(* IEC 61131-3 sources: daoli-st-library/DL_Algo (part 12) *)

(* ---- FB_DL_EtchEndpointTrend.st ---- *)
(*==============================================================================
 * 组件名称 (Component)  : FB_DL_EtchEndpointTrend
 * 所属子库 (Sublibrary) : DL_Algo
 * 前缀     (Prefix)     : FB_DL_
 * 当前版本 (Version)    : 1.0.1
 * 兼容性   (Platform)   : CODESYS 3.5 / TwinCAT 3 / 汇川 InoProShop / Schneider
 *                         Machine Expert；纯 IEC 61131-3（第 3 版），
 *                         仅依赖标准库 TON / ABS / MAX / MIN 与库内
 *                         FB_DL_Differentiator（IN-OUT 注入消费），
 *                         零厂商方言
 * 作者     (Author)     : 道莅代码库 · PLC编程专家（R31）
 * 开源溯源 (Origin)     : 刻蚀终点趋势检测公开工艺语义（行业池主源；
 *                         Measurement 行统计族语义邻接不重复记账），道莅
 *                         clean-room 防御性实现，未复制任何外部源码行
 * 功能描述 (Function)   : 刻蚀终点趋势双判据检测件。学习相采基线（均值与
 *                         噪声窗）；监视相用库内 FB_DL_Differentiator 求变化
 *                         率（IN-OUT 注入，不内联），斜率换算为 单位每分钟；
 *                         双判据：斜率绝对值超阈 且 信号突破噪声窗，持续
 *                         tConf 触发终点并锁存，保持至 bRun 下降显式复位。
 *                         斜率量纲占位说明：fSignal 的工程单位由调用方定义，
 *                         fSlope 与 fSlopeTh 同量纲，单位为 调用方单位每分钟。
 * 依赖表   (Depends)    : FB_DL_Differentiator（微分器，IN-OUT 注入消费，
 *                         本件不内联差分）。
 * 状态机   (States)     : eLearning/eMonitor/eTriggered，CASE 带 ELSE 复位
 *                         回学习相（信息级提示）。
 * 码位     (Codes)      : 16#0002_3033 信息级：信号非有限冻结评估、学习相
 *                                      非有限重启学习、样本不足不出判定
 *                                      （不置 bError）
 *                         16#0002_3034 故障级：确认窗中断判据矛盾（锁存）
 *                         16#0002_3035~0037 保留未启用（码表与实现对齐）
 * 边界防错 (Boundary)   : 1 信号非有限（x<>x 自反判加幅值界）监视相冻结评估、
 *                           学习相清积累重启学习；
 *                         2 学习相样本不足不出判定；
 *                         3 斜率时间差防除零由库内微分器公共钳位承担
 *                           （其 fDt 下限 10 毫秒），本件不做二次除法；
 *                         4 TON 实例每拍无条件刷新；
 *                         5 触发锁存可达解除路径：bRun 下降沿显式复位；
 *                         6 确认窗中途判据消失按判据矛盾锁故障。
 * 修订历史 (Revision)   : 2026-11-18 v1.0.0 首版入库（R31 · 阶段三 · 序 20）
 *                         2026-11-18 v1.0.1 R31 终审修复：先验基线模式补
 *                         uCnt 计数，消除方差分母 1E-30 退化致判据二永假
 *==============================================================================*)

(*------------------------------------------------------------------------------
 * 枚举: E_DL_EndpointState（归属本功能块，同文件发布，全库唯一属主）
 *----------------------------------------------------------------------------*)
TYPE E_DL_EndpointState :
(
    eLearning  := 0,   // 学习相：采基线均值与噪声窗 / Learning, baseline mean and noise window
    eMonitor   := 10,  // 监视相：双判据评估 / Monitor, dual-criteria evaluation
    eTriggered := 20   // 触发相：终点锁存至显式复位 / Triggered, endpoint latched until explicit reset
);
END_TYPE

(*==============================================================================
 * 功能块: FB_DL_EtchEndpointTrend
 * 调用约定: 每个扫描周期无条件调用一次；ioDiff 为调用方持有的库内微分器
 *           实例（IN-OUT 注入），本件驱动其引脚并读取其输出。
 *==============================================================================*)
FUNCTION_BLOCK FB_DL_EtchEndpointTrend
VAR_INPUT
    fSignal   : LREAL := 0.0;         // 工艺信号 [调用方单位] / Process signal [caller unit]
    bRun      : BOOL := FALSE;        // 工步运行（下降沿显式复位）/ Process running, falling edge resets
    fSlopeTh  : REAL := 5.0;          // 斜率判据阈 [调用方单位每分钟] / Slope threshold [caller unit per min]
    fNoiseWin : REAL := 2.0;          // 噪声窗 [调用方单位] / Noise window [caller unit]
    tConf     : TIME := T#3S;         // 触发确认窗时长 [毫秒] / Trigger confirm window [ms]
    fBaseline : LREAL := 0.0;         // 外部先验基线（0 = 无先验走自采）/ External prior baseline, 0 = none
    tLearn    : TIME := T#30S;        // 学习相时长 [毫秒]（可增引脚）/ Learning duration [ms], added pin
    tSample   : TIME := T#500MS;      // 微分器采样周期 [毫秒]（可增引脚）/ Differentiator sample period [ms], added pin
END_VAR
VAR_IN_OUT
    ioDiff    : FB_DL_Differentiator; // 库内微分器实例注入（斜率不内联）/ Library differentiator instance injected
END_VAR
VAR_OUTPUT
    bEndpoint : BOOL;                 // 终点触发锁存输出 / Endpoint trigger latched output
    fSlope    : REAL;                 // 斜率输出 [调用方单位每分钟] / Slope output [caller unit per min]
    eState    : E_DL_EndpointState;   // 判定状态 / Detection state
    bError    : BOOL;                 // 故障标志，与故障级码配对（R45）/ Fault flag paired with fault codes
    uErrorId  : UDINT;                // 错误码，0 = 无错 / Error code, 0 = none
END_VAR
VAR
    tonLearn  : TON;                  // 学习相计时，每拍无条件刷新 / Learning timer, refreshed every scan
    tonConf   : TON;                  // 触发确认窗计时，每拍无条件刷新 / Confirm window timer, refreshed every scan
    fSigR     : REAL;                 // 信号 REAL 域副本 [调用方单位] / Signal REAL copy [caller unit]
    bSigOk    : BOOL;                 // 信号有限有效 / Signal finiteness validity
    fSum      : REAL;                 // 学习相样本和 [调用方单位] / Learning sample sum [caller unit]
    fSumSq    : REAL;                 // 学习相平方和 [平方调用方单位] / Learning sum of squares
    uCnt      : UDINT;                // 学习相样本数 [个] / Learning sample count
    fMean     : REAL;                 // 基线均值 [调用方单位] / Baseline mean [caller unit]
    fNoise    : REAL;                 // 噪声窗实测 [调用方单位] / Measured noise window [caller unit]
    bLearnDone: BOOL;                 // 学习完成标志 / Learning done flag
    bCritSlope: BOOL;                 // 判据一：斜率超阈 / Criterion one, slope over threshold
    bCritNoise: BOOL;                 // 判据二：突破噪声窗 / Criterion two, beyond noise window
    bCritNow  : BOOL;                 // 双判据本拍合取 / Both criteria this scan
    bInWin    : BOOL;                 // 确认窗进行中 / Confirm window in progress
    bPriorUse : BOOL;                 // 先验基线使用标志 / Prior baseline usage flag
    uCodeLatch: UDINT;                // 故障级锁存码 / Latched fault code
END_VAR
VAR CONSTANT
    DL_EET_FIN   : LREAL := 1.0E30;   // LREAL 有限幅值判界 / LREAL finiteness magnitude bound
    DL_EET_FINR  : REAL  := 1.0E30;   // REAL 有限幅值判界 / REAL finiteness magnitude bound
    DL_EET_MIN   : UDINT := 20;       // 学习相最少样本数 [个] / Learning minimum samples
    DL_EET_MIN60 : REAL  := 60.0;     // 每秒到每分钟换算系数 / Per-second to per-minute factor
    DL_EET_EPS   : REAL  := 1.0E-30;  // 样本数防除零容差 / Sample count divide guard
END_VAR

// ---- 段 1｜定时器实例无条件周期刷新（红线：禁入条件分支）----------------------
tonLearn(IN := (eState = eLearning) AND bRun, PT := tLearn);   // 学习计时 / Learning timing
tonConf(IN := bCritNow, PT := tConf);                          // 确认窗计时无条件 / Confirm timing unconditionally

// ---- 段 2｜信号有效性（自反判加幅值界）----------------------------------------
bSigOk := (fSignal = fSignal) AND (ABS(fSignal) < DL_EET_FIN); // 信号有限 / Signal finite
fSigR := LREAL_TO_REAL(fSignal);                               // 信号落 REAL 域 / Signal to REAL domain

// ---- 段 3｜显式复位：bRun 下降沿清全部锁存 ------------------------------------
IF NOT bRun THEN
    bEndpoint := FALSE;                            // 复位清终点锁存 / Reset clears endpoint latch
    IF eState = eTriggered THEN
        eState := eLearning;                       // 触发相复位回学习 / Triggered resets to learning
    END_IF
END_IF

// ---- 段 4｜驱动库内微分器（IN-OUT 注入，输出即变化率 单位每秒）----------------
ioDiff(bEnable := bRun AND bSigOk,                    // 信号无效停微分防伪速率 / Invalid signal stops differentiator
       fIn := fSigR,                                  // 被微分量注入 / Differentiated input injected
       tFiltTime := T#1S,                             // 低通时间常数固定档 / Fixed low-pass constant
       tSampleTime := tSample);                       // 采样周期透传 / Sample period passed
fSlope := ioDiff.fRateOut * DL_EET_MIN60;             // 斜率换算每分钟（量纲占位见头注释）/ Slope per minute

// ---- 段 5｜学习相：采基线均值与噪声窗 ------------------------------------------
IF (eState = eLearning) AND bRun THEN
    IF NOT bSigOk THEN
        fSum := 0.0;                                  // 非有限清积累重启学习（信息级）/ Non-finite restarts learning
        fSumSq := 0.0;                                // 清平方和积累 / Clear sum-of-squares
        uCnt := 0;                                    // 清样本计数 / Clear sample count
        bLearnDone := FALSE;                          // 撤完成标志 / Withdraw done flag
        uErrorId := 16#0002_3033;                     // 信息级：学习重启 / Info: learning restarted
    ELSE
        bPriorUse := (fBaseline <> 0.0) AND (fBaseline = fBaseline)
                 AND (ABS(fBaseline) < DL_EET_FIN);   // 先验基线可用性 / Prior baseline availability
        IF bPriorUse THEN
            fMean := LREAL_TO_REAL(fBaseline);        // 先验均值直接生效 / Prior mean applied directly
            uCnt := uCnt + 1;                         // 先验模式同样计数（方差分母防爆，R28 终审）/ Prior mode counts samples too
        ELSE
            fSum := fSum + fSigR;                     // 自采样本累加 / Self-sample accumulation
            uCnt := uCnt + 1;                         // 样本计数 / Sample count
        END_IF
        fSumSq := fSumSq + fSigR * fSigR;             // 平方和积累（样本方差用）/ Sum of squares accumulation
        IF tonLearn.Q AND (bPriorUse OR (uCnt >= DL_EET_MIN)) THEN
            IF NOT bPriorUse THEN
                fMean := fSum / UDINT_TO_REAL(uCnt);  // 均值收口，分母已验下限 / Mean closed, denominator verified
            END_IF
            fNoise := SQRT(MAX(fSumSq / MAX(UDINT_TO_REAL(uCnt), DL_EET_EPS) - fMean * fMean, 0.0)); // 样本标准差收口（平方和法）/ Sample stddev via sum-of-squares
            bLearnDone := TRUE;                       // 学习完成 / Learning done
            eState := eMonitor;                       // 转监视相 / To monitor
        END_IF
    END_IF
END_IF

// ---- 段 6｜监视相：双判据评估与确认窗 ------------------------------------------
IF (eState = eMonitor) AND bRun THEN
    IF NOT bSigOk OR (NOT ioDiff.bValid) THEN
        bCritSlope := FALSE;                          // 数据无效撤判据一 / Invalid data withdraws criterion one
        bCritNoise := FALSE;                          // 数据无效撤判据二 / Invalid data withdraws criterion two
        uErrorId := 16#0002_3033;                     // 信息级：冻结评估 / Info: evaluation frozen
    ELSIF (uCnt < DL_EET_MIN) AND (NOT bPriorUse) THEN
        bCritSlope := FALSE;                          // 样本不足不出判定 / Insufficient samples, no verdict
        bCritNoise := FALSE;                          // 样本不足不出判定 / Insufficient samples, no verdict
        uErrorId := 16#0002_3033;                     // 信息级：样本不足 / Info: insufficient samples
    ELSE
        bCritSlope := ABS(fSlope) > ABS(fSlopeTh);    // 判据一：斜率超阈 / Slope over threshold
        bCritNoise := ABS(fSigR - fMean) > fNoise;    // 判据二：突破噪声窗 / Beyond noise window
    END_IF
    bCritNow := bCritSlope AND bCritNoise;            // 双判据合取 / Both criteria AND
    bInWin := (tonConf.ET > T#0MS);                   // 确认窗进行中判定 / Confirm window in progress
    IF bInWin AND (NOT bCritNow) THEN
        eState := eLearning;                          // 按判据矛盾复位回学习重采基线 / Contradiction resets to learning
        uCodeLatch := 16#0002_3034;                   // 码位：确认窗中断判据矛盾 / Code: confirm window contradiction
        bError := TRUE;                               // 故障级配对置位（R45）/ Fault flag paired
    ELSIF tonConf.Q THEN
        bEndpoint := TRUE;                            // 确认满终点触发锁存 / Confirmed, endpoint latched
        eState := eTriggered;                         // 转触发相 / To triggered
        bError := FALSE;                              // 清故障标志 / Clear fault flag
        uCodeLatch := 16#0000_0000;                   // 清锁存码 / Clear latched code
    END_IF
END_IF

// ---- 段 7｜错误码装配：故障锁存回放优先，信息级居次 -----------------------------
IF (eState = eLearning) AND bRun AND (uCodeLatch <> 16#0000_0000) THEN
    bError := TRUE;                                   // 故障锁存回放（学习相等待重试）/ Fault latched replay
    uErrorId := uCodeLatch;                           // 锁存码回放 / Latched code replayed
ELSIF NOT bRun THEN
    bError := FALSE;                                  // 撤运行清故障（可达解除）/ Run drop clears fault
    uErrorId := 16#0000_0000;                         // 清码 / Clear code
    uCodeLatch := 16#0000_0000;                       // 清锁存码 / Clear latched code
END_IF
END_FUNCTION_BLOCK

(* ---- FB_DL_EwmaFilter.st ---- *)
(*
  ==================================================================
  组件名 Component  : FB_DL_EwmaFilter
  分类   Category   : DL_Algo
  前缀   Naming     : FB_DL_ ｜ b/n/u/f/t/e/st 类型前缀制（R265）
  码位   Code ID    : 16#0002_373B / 373C（故障级）
  版本   Version    : 1.0.0
  复杂度 Complexity  : 低
  功能   Purpose    : EWMA 指数加权滑动平均 fOut := fOut + α×(fIn − fOut)，α 直接
                      入参（离散统计 / SPC 平滑口径），供调用方直接整定平滑系数。
  开源溯源 Origin    : 公开公式 clean-room，参考公开统计过程控制（SPC）教材的
                      EWMA 定义（分类与公式借鉴，零代码复制），本件实现、闸门与
                      码位 100% 自有。
  许可证 License    : MIT
  参考   Reference  : IEC 61131-3:2013 §6.6 算术运算符；EWMA 递推式 y[k] =
                      y[k−1] + α·(x[k] − y[k−1]) 为公开统计公式
  平台   Platform   : 纯 IEC 61131-3（四则 / 比较），三平台通用
  依赖   Depends    : 仅 Standard.library（无库调用、无定时器）
  分工声明 Split     : FB_DL_LowPassFilter 为连续时间常数口径（α 由 tTf / tDt 派生，
                      一阶 RC 语义）；FB_DL_MovingAverage 为等权滑窗；本件为调用方
                      直接给 α 的统计平滑口径（EWMA / SPC 语义）；三者选型对照进
                      MANUAL_DL_Algo（R216 双向互引）。
  归属 Ownership     : 本件无 TYPE 声明；全部引脚为 IEC 标准原生类型。
  ------------------------------------------------------------------
  边界 Boundary     :
                      一 α 域闸 (0, 1]：fAlpha <= 0 或 > 1 或非有限 → 组态码 373B +
                         出口三件套 + RETURN 结构早退（开区间下界防输出冻结，
                         α = 0 是「禁冻结伪装正常」的组态错误而非合法参数）；
                      二 fIn 非有限（NaN / ±Inf）→ 本拍拒绝更新、保持上拍有效值 +
                         故障码 373C + 三件套（禁污染物进入递推状态）；
                      三 首拍 _bInit → fOut := fIn 首样本直通（禁输出 0 假跳变）；
                      四 bEnable = FALSE 的语义写死（FB33-4 声明行）：本件取「冻结
                         最后有效值」，理由：纯监视滤波不驱动功率级，冻结均值供
                         HMI 连续读数（与 BiquadFilter 的「控制量归零」口径不同，
                         选型时注意）；
                      五 故障码策略（本件无 bReset 引脚，R152 解除路径自证）：组态类
                         与测量类故障码逐拍重算不锁存，解除路径 = 修正组态 / 恢复
                         测点（恒可达）；首因保序由判据顺序保证；
                      六 非有限闸逐个点名（R272）：fAlpha 与 fIn 双双入闸；
                      七 首拍 _bInit 全量初始化（FB50-2）；无定时器 / 无边沿实例，
                         段 0 无刷新对象（R6 标注 N/A）；无全局、无外部变量、无
                         物理地址、无指针。
  错误码 Codes      :
    16#0002_373B【故障级】组态非法（fAlpha ≤ 0 / > 1 / 非有限）
    16#0002_373C【故障级】输入非有限（fIn 为 NaN / ±Inf）或递推结果非有限（后者
                         理论上不可达的兜底分支，与输入坏同码，出口组合不可区分，
                         R90 反证：fOut 保持上拍有效值 + bValid = FALSE 两场景同形）
  码位反证 Note     :
    373B 与 373C 不可合并：两者的处置人不同（组态工程师调 α / 仪表工查测点），
    而两者出口组合不同（组态坏无论 fIn 有限与否恒发 373B），可由场景唯一还原，
    故分立两码（R90）。
  验收 Acceptance   :
    算法已证（脚本）：未跑 ｜ 编译器已证（三平台）：未跑
    V1 α = 1 → 直通 fOut = fIn（逐拍断言）
    V2 α = 0 → 码 373B + 三件套 + 早退（禁冻结伪装正常）
    V3 α = 0.5 阶跃 0 → 100 → 逐拍 50 / 75 / 87.5 收敛，无超调
    V4 fIn = NaN → 保持上拍 fOut + 码 373C + bValid = FALSE
    V5 首拍 → fOut = fIn 首样本直通（禁 0 假跳变）
    V6 bEnable = FALSE → fOut 冻结最后有效值（边界四声明行回归向量）
  修订记录 Revision  :
    2026-11-21  v1.0.0  R63 首版（批 1 · 序号 3）
  ==================================================================
*)
FUNCTION_BLOCK FB_DL_EwmaFilter
VAR_INPUT
    bEnable  : BOOL := TRUE;  // 使能，FALSE 时输出冻结最后有效值（边界四）/ the enable, false freezes the last valid output
    fIn      : LREAL := 0.0;  // 输入量 [工程单位]，必须有限 / the input value, must be finite
    fAlpha   : LREAL := 0.2;  // 平滑系数 [−]，合法域 (0, 1] 开区间下界 / the smoothing factor inside the half open domain from zero exclusive to one
END_VAR
VAR_OUTPUT
    fOut     : LREAL := 0.0;           // 滤波输出 [工程单位] / the filtered output
    bValid   : BOOL := FALSE;          // 输出可用（使能 + 无故障 + 首样本已收）[-] / the output is usable
    eErr     : UDINT := 16#0000_0000;  // 错误码，0 = 正常 / the error code, zero is ok
    bError   : BOOL := FALSE;          // 故障标志（故障级码同拍置位，R45 配对）/ the fault flag raised with a fault level code
END_VAR
VAR
    _bInit    : BOOL := FALSE;   // 首拍初始化标志（R310 / FB50-2）/ the first scan flag
    _bHasSamp : BOOL := FALSE;   // 已收首样本标志（跨拍保持）/ the first sample received flag
    _fOutLast : LREAL := 0.0;    // 最近一次有效输出（冻结与递推基线）[工程单位] / the last valid output used as the freeze and the recursion base
    _bFinIn   : BOOL := FALSE;   // 输入有限闸结果（逐拍重算）/ the input finiteness gate result
    _bFinAlp  : BOOL := FALSE;   // 平滑系数有限闸结果（逐拍重算）/ the alpha finiteness gate result
END_VAR  // R64 结构补齐：VAR 段缺失的 END_VAR（门禁机械修复）
VAR CONSTANT
    DL_EWM_ZERO : LREAL := 0.0; // 实数零常量 [工程单位] / the real zero constant
    DL_EWM_ONE  : LREAL := 1.0; // 实数一常量（α 上界）[-] / the real unit constant, the alpha ceiling
END_VAR

// 段 0｜本件无定时器与边沿实例（纯递推滤波器，R6 标注 N/A），无刷新对象 / segment 0, no timers and no edge instances exist here

// 段 1｜首拍初始化（FB50-2）/ segment 1, the first scan init
IF NOT _bInit THEN // 首拍一拍 / the first scan
    _bInit := TRUE; // 置首拍标志 / raise the first scan flag
    _bHasSamp := FALSE; // 首样本标志显式清零（触发首拍直通）/ clear the first sample flag so the direct pass triggers
    _fOutLast := DL_EWM_ZERO; // 最近有效输出显式清零 / clear the last valid output explicitly
END_IF

// 段 2｜非有限闸逐个点名（R272：fAlpha 与 fIn 双双入闸）/ segment 2, the finiteness gates naming both real pins
_bFinAlp := (fAlpha = fAlpha) AND ((fAlpha - fAlpha) = (fAlpha - fAlpha)); // 平滑系数有限 / the alpha is finite
_bFinIn := (fIn = fIn) AND ((fIn - fIn) = (fIn - fIn)); // 输入有限 / the input is finite

// 段 3｜α 组态域闸：结构早退（边界一，出口三件套 + RETURN）/ segment 3, the alpha domain gate with the structural early exit
IF (NOT _bFinAlp) OR (fAlpha <= DL_EWM_ZERO) OR (fAlpha > DL_EWM_ONE) THEN // 组态非法 / an illegal configuration
    fOut := _fOutLast; // 出口保持最近有效值（禁自赋值出口，R261）/ keep the last valid output instead of a self assignment
    bValid := FALSE; // 输出不可用 / the output is not usable
    eErr := 16#0002_373B; // 故障级：α 组态非法 / fault grade, the alpha configuration is illegal
    bError := TRUE; // 同拍置故障标志（R45 配对）/ raise the fault flag on the same scan
    RETURN; // 早退（组态非法结构早退，R1 同族口径）/ early return, the structural exit on an illegal configuration
END_IF

// 段 4｜失能分支：冻结最后有效值（边界四声明行）/ segment 4, the disabled branch freezes the last valid output
IF NOT bEnable THEN // 失能 / disabled
    fOut := _fOutLast; // 冻结最后有效值（纯监视滤波，理由见边界四）/ freeze the last valid output, a pure monitoring filter
    bValid := FALSE; // 失能即不可用 / the output is not usable while disabled
    bError := FALSE; // 失能不是故障 / a disabled device is not a fault
    eErr := 16#0000_0000; // 失能不发码 / no code is emitted while disabled
    RETURN; // 早退，不推进递推 / early return without advancing the recursion
END_IF

// 段 5｜输入非有限：拒绝更新并保持（边界二，禁污染物进状态）/ segment 5, a non finite input is rejected
IF NOT _bFinIn THEN // 输入坏 / the input is broken
    fOut := _fOutLast; // 保持上拍有效值 [工程单位] / keep the last valid output
    bValid := FALSE; // 输出不可用 / the output is not usable
    eErr := 16#0002_373C; // 故障级：输入非有限 / fault grade, the input is not finite
    bError := TRUE; // 同拍置故障标志（R45 配对）/ raise the fault flag on the same scan
    RETURN; // 早退，递推状态不被污染 / early return, the recursion state stays clean
END_IF

// 段 6｜首样本直通（边界三，禁 0 假跳变）/ segment 6, the first sample passes straight through
IF NOT _bHasSamp THEN // 尚无首样本 / no first sample yet
    _fOutLast := fIn; // 基线 = 首样本 [工程单位] / the base is the first sample
    _bHasSamp := TRUE; // 置首样本标志 / raise the first sample flag
    fOut := fIn; // 首拍直通 [工程单位] / the first scan passes straight through
    bValid := TRUE; // 输出可用 / the output is usable
    eErr := 16#0000_0000; // 正常 / ok
    bError := FALSE; // 无故障 / no fault
    RETURN; // 早退 / early return
END_IF

// 段 7｜EWMA 递推（公开公式）：fOut = fOutLast + α×(fIn − fOutLast) / segment 7, the EWMA recursion
fOut := _fOutLast + (fAlpha * (fIn - _fOutLast)); // 指数加权滑动平均 [工程单位] / the exponentially weighted moving average

// 段 8｜递推结果非有限兜底（三件套，R258；与输入坏同码，反证见码表）/ segment 8, the non finite result fallback
IF (fOut <> fOut) OR ((fOut - fOut) <> (fOut - fOut)) THEN // 结果非有限（NaN 自反 / Inf 差值自减）/ a non finite result tested by reflexivity and the self difference
    fOut := _fOutLast; // 回退保持上拍有效值 [工程单位] / fall back to the last valid output
    bValid := FALSE; // 输出不可用 / the output is not usable
    eErr := 16#0002_373C; // 故障级：输入或结果非有限（同族一码）/ fault grade, the input or the result is not finite
    bError := TRUE; // 同拍置故障标志（R45 配对）/ raise the fault flag on the same scan
    RETURN; // 早退，基线不被污染 / early return, the base stays clean
END_IF

// 段 9｜统一出口（基线推进 + 可用声明）/ segment 9, the unified outlet
_fOutLast := fOut; // 基线推进（写前已过非有限闸）[工程单位] / advance the base after the finiteness gate
bValid := TRUE; // 输出可用 / the output is usable
bError := FALSE; // 无故障 / no fault
eErr := 16#0000_0000; // 正常 / ok
END_FUNCTION_BLOCK

(* ---- FB_DL_ExcessAirTrim.st ---- *)
(*==============================================================================
 * 组件名称 (Component)  : FB_DL_ExcessAirTrim
 * 溯源说明 (Provenance): 道莅 clean-room 防御性实现（IEC 61131-3 纯净实现，闭源文档仅借语义，零代码行）
 * 所属子库 (Sublibrary) : DL_Algo / ProcessControl
 * 当前版本 (Version)    : 1.0.0
 * 兼容性   (Platform)   : CODESYS 3.5 / TwinCAT 3 / 汇川 InoProShop / 施耐德
 *                         Machine Expert；纯 IEC 61131-3（第 3 版），仅用
 *                         Standard.library 的 TON / LIMIT / ABS / TIME_TO_DINT / DINT_TO_TIME
 * 组件分类 (Category)   : 功能块（FUNCTION_BLOCK）· 氧量修正（空燃比长期偏置）
 * 功能一句话 (Summary)  : 按烟气含氧量与目标的偏差，按固定步长缓慢修正空燃比，
 *                         越死区才动、负荷剧变时冻结、修正量双侧钳位。
 *
 * 本件存在的意义 (Why this unit exists)
 *   与 FB_DL_CrossLimitSelect 是互补的两条律：交叉限幅管「同拍谁先给」，
 *   本件管「长期空燃比偏置」。二者不可合并——一个是逐拍代数选择，
 *   一个是慢时标步进律，合并后验收向量无法独立手算复算。
 *   ROADMAP §7 的锅炉/加热炉条目全部依赖这一对。
 *
 * 时间标度 (Time scale)
 *   步进节拍 = tConfirm：偏差持续 tConfirm 才走一步 fTrimStep。因此修正速率
 *   ≈ fTrimStep / tConfirm（例：0.05 % / 30 s ≈ 0.1 %/min），比燃烧回路慢两到
 *   三个数量级——这是刻意的：氧量探头本身有分钟级滞后，快修正只会来回过冲。
 *   tConfirm = T#0S 是合法语义（每拍一步），不置错，但此时步进率与扫描周期绑定，
 *   属调用方自担的用法，已在此声明。
 *
 * 边界安全 (Boundary)
 *   ① fO2Target <= 0、fO2Deadband < 0、fTrimLimit <= 0、fTrimStep <= 0，或四者
 *      任一非有限 → 故障 2C10，fTrim := 0（退回纯交叉限幅，安全可利用）；
 *   ② 氧量或负荷率非有限 → 故障 2C11，**保持末次 fTrim**（坏值不得清掉长期偏置）；
 *   ③ 死区内 → 信息 2C01，不修正、fTrim 保持；
 *   ④ |fLoadRate| > fRateFreeze → 信息 2C02，冻结修正、fTrim 保持；
 *   ⑤ 累加后双侧钳 ±fTrimLimit（抗饱和，不做积分回算）；
 *   ⑥ 失能 → eIdle，fTrim := 0 且**保持量一并清 0**，避免再使能时旧偏置
 *      突然回投（无扰投切，见 FB_DL_ExcessAirTrim 组装说明）；
 *   ⑦ TON 实例在主体最前部无条件刷新，步进后经「断输入一拍」标志重启计时，
 *      使步进节拍严格等于 tConfirm；
 *   ⑧ CASE 落 ELSE 置 2C12 并回 eFault。
 *
 * 错误码    : 16#0002_2C01 偏差在死区内，不修正（fTrim 保持）——信息级，正常调节
 *             16#0002_2C02 负荷变化率超限，修正已冻结——信息级，保护动作
 *             16#0002_2C10 修正参数非法（目标/死区/限幅/步长），fTrim 归零——故障级
 *             16#0002_2C11 氧量或负荷率非有限，保持末次 fTrim——故障级
 *             16#0002_2C12 状态机落 ELSE 兜底（非法状态）——故障级，回 eFault
 * 码位总账  : 16#0002_2C01 用 / 16#0002_2C02 用 ｜ 16#0002_2C10 用 / 16#0002_2C11 用 / 16#0002_2C12 用
 * 状态机    : E_DL_O2TrimState（eIdle / eActive / eFrozen / eFault），CASE 含 ELSE 兜底，
 *             ELSE 置 16#0002_2C12 并回 eFault；失能无条件回 eIdle
 * 采样约定  : 每任务周期调用一次；修正节拍由 tConfirm 决定，不读系统时钟
 * 依赖说明  : 零 DL_ 子库依赖（DL_Algo 只允许 Standard.library，限幅与死区内联实现）
 * 验收向量  : V1 氧量 4.0 %、目标 3.0 %、死区 0.3、tConfirm 30 s → 每 30 s 走一步
 *               fTrim −0.05，单调减到 −5.0 后钳住（抗饱和主向量）
 *             V2 氧量 3.2 %（死区内）→ 不修正，eErr = 2C01，fTrim 不动
 *             V3 fLoadRate = 5 %/s > fRateFreeze → bFrozen = TRUE，eErr = 2C02，fTrim 不动
 *             V4 fO2Target = 0 → fTrim = 0，eErr = 2C10，bError = TRUE，eFault
 *             V5 fO2Meas = NaN → fTrim 保持上一拍值，eErr = 2C11（保持主向量）
 *             V6 bEnable 落 → eIdle，fTrim = 0、bActive = FALSE、保持量清 0（恢复首拍不阶跃）
 *             V7 tConfirm = T#0S → 每拍一步，不置错（合法语义向量）
 * 红线自检  : 全局变量声明零使用 / 外部变量访问零使用 / 物理地址零使用 ｜ 纯 IEC 61131-3 ｜ 除法仅一处
 *             常量除（无除零面）｜ 浮点只用大小与容差比较 ｜ 无循环 ｜ 全变量双语
 *             同行注释 ｜ ENUM + CASE 含 ELSE ｜ TON 在主体最前部无条件刷新 ｜
 *             无魔法数
 * 修订历史  : 2026-11-16  v1.0.0  首版入库（R22 · 批 2 · 燃烧保护律）
 *============================================================================*)

(*-----------------------------------------------------------------------------
 * 枚举: E_DL_O2TrimState（归属本功能块，同文件发布，全库唯一定义）
 * 含义: 氧量修正的工作相位。0 起步长 10。
 *-----------------------------------------------------------------------------*)
TYPE E_DL_O2TrimState :
(
    eIdle    := 0,     // 待机：未使能或参数非法，修正量为 0 / Idle, disabled or illegal parameters, trim is zero
    eActive  := 10,    // 生效：越死区且负荷平稳，按节拍步进 / Active, outside the dead band with a steady load
    eFrozen  := 20,    // 冻结：负荷变化率超限，保持修正 / Frozen, load rate above the limit, trim held
    eFault   := 99     // 故障：参数非法或输入非有限 / Fault, illegal parameter or non-finite input
);
END_TYPE

FUNCTION_BLOCK FB_DL_ExcessAirTrim
VAR_INPUT
    fO2Meas      : REAL;                       // 烟气含氧量实测 [%]，范围 0~21 / measured flue gas oxygen [%], range 0~21
    fO2Target    : REAL := 3.0;                // 目标氧含量 [%]，须 > 0 / target oxygen content [%], must be > 0
    fO2Deadband  : REAL := 0.3;                // 死区半宽 [%]，须 >= 0 / dead band half width [%], must be >= 0
    fTrimLimit   : REAL := 5.0;                // 修正量上限 [%]，对称，须 > 0 / symmetric trim limit [%], must be > 0
    fTrimStep    : REAL := 0.05;               // 单步修正量 [%]，须 > 0 / single trim step [%], must be > 0
    fLoadRate    : REAL;                       // 负荷变化率 [%/s] / load change rate [%/s]
    fRateFreeze  : REAL := 2.0;                // 冻结门限 [%/s]，须 > 0 / freeze threshold [%/s], must be > 0
    tConfirm     : TIME := T#30S;              // 步进确认时间 [ms]，0 = 每拍一步 / step confirm time [ms], zero means one step per scan
    bEnable      : BOOL;                       // 使能 / enable
END_VAR
VAR_OUTPUT
    fTrim        : REAL;                       // 空燃比修正量 [%]，正为增空气 / air to fuel ratio trim [%], positive adds air
    bActive      : BOOL;                       // 修正生效标志 / trim active flag
    bFrozen      : BOOL;                       // 修正冻结标志 / trim frozen flag
    eErr         : UDINT;                      // 错误码，0 表示无错 / error code, 0 means no error
    bError       : BOOL;                       // 故障级标志，仅故障级错误置位 / fault-class flag, set only on fault-level codes
    bValid       : BOOL;                       // 输出可用标志 / outputs usable flag
END_VAR
VAR
    fbConfirm    : TON;                        // 步进节拍计时，段 5 无条件刷新 [ms] / step cadence timer, refreshed unconditionally
    _eState      : E_DL_O2TrimState := E_DL_O2TrimState.eIdle; // 当前相位 / current phase
    _bInit       : BOOL := FALSE;              // 首扫标志，初值 FALSE 取非判定 / first-scan flag, tested negated
    _bParamBad   : BOOL;                       // 参数非法标志 / illegal parameter flag
    _bFiniteBad  : BOOL;                       // 输入非有限标志 / non-finite input flag
    _bIllegal    : BOOL;                       // 非法状态标志 / illegal state flag
    _bCond       : BOOL;                       // 步进条件（越死区且负荷平稳） / step condition, outside dead band with a steady load
    _bStepPulse  : BOOL;                       // 本拍步进脉冲 / step pulse of this scan
    _bConfirmBreak : BOOL;                     // 节拍计时器断输入一拍标志 / cadence timer one-scan break flag
    _tConfirmUse : TIME := T#30S;              // 生效确认时间 [ms]，已钳位 / effective confirm time, clamped
    _fTrimHeld   : REAL;                       // 修正量保持量 [%] / held trim [%]
    _fDev        : REAL;                       // 氧量偏差 = 实测 − 目标 [%] / oxygen deviation, measured minus target
    _fAbsDev     : REAL;                       // 偏差绝对值 [%] / absolute deviation [%]
    _fAbsRate    : REAL;                       // 负荷变化率绝对值 [%/s] / absolute load rate [%/s]
    _fBandUse    : REAL := 0.3;                // 生效死区半宽 [%] / effective dead band half width
END_VAR
VAR CONSTANT
    DL_VAL_LIM   : REAL := 1.0E30;             // 有限性判定的绝对值上限 [无量纲] / finiteness ceiling
    DL_O2_MAX    : REAL := 21.0;               // 氧量物理上限 [%] / physical oxygen ceiling [%]
    DL_TARGET_MN : REAL := 0.0;                // 目标氧含量下限 [%]，须严格大于 / target oxygen floor, must be strictly greater
    DL_BAND_MN   : REAL := 0.0;                // 死区半宽下限 [%] / dead band floor [%]
    DL_LIMIT_MN  : REAL := 0.0;                // 修正限幅下限 [%]，须严格大于 / trim limit floor, must be strictly greater
    DL_STEP_MN   : REAL := 0.0;                // 步长下限 [%]，须严格大于 / step floor, must be strictly greater
    DL_RATE_MN   : REAL := 0.0;                // 冻结门限下限 [%/s]，须严格大于 / freeze threshold floor, must be strictly greater
    DL_EPS       : REAL := 1.0E-6;             // 浮点比较容差 [%] / float comparison tolerance [%]
    DL_CONF_MAX_MS : DINT := 3600000;          // 确认时间上限 [ms]，一小时 / confirm time ceiling, one hour
    DL_TIME_ZERO : TIME := T#0MS;              // 时间零值基准 [ms] / time zero reference
END_VAR

(*------------------------------------------------------------------------------
 * 段 1｜每拍预置（保持量与输出在段 8 单点写入，此处不清）
 *      Per-scan presets, held values and outputs are written only in segment eight
 *-----------------------------------------------------------------------------*)
eErr        := 16#0000_0000;                   // 错误码每拍重算 / error code recomputed every scan
bError      := FALSE;                          // 故障标志每拍重算 / fault flag recomputed every scan
bValid      := FALSE;                          // 可用标志每拍重算 / usable flag recomputed every scan
bActive     := FALSE;                          // 生效标志每拍重算 / active flag recomputed every scan
bFrozen     := FALSE;                          // 冻结标志每拍重算 / frozen flag recomputed every scan
_bParamBad  := FALSE;                          // 参数非法标志预清零 / parameter flag pre-cleared
_bFiniteBad := FALSE;                          // 非有限标志预清零 / non-finite flag pre-cleared
_bIllegal   := FALSE;                          // 非法状态标志预清零 / illegal state flag pre-cleared
_bCond      := FALSE;                          // 步进条件预置 FALSE / step condition preset FALSE
_bStepPulse := FALSE;                          // 步进脉冲预置 FALSE / step pulse preset FALSE

(*------------------------------------------------------------------------------
 * 段 2｜首扫初始化（修正量从 0 起：投用即无偏置，符合无扰投切）
 *      First-scan initialisation, the trim starts at zero for a bumpless start
 *-----------------------------------------------------------------------------*)
IF NOT _bInit THEN
    _eState      := E_DL_O2TrimState.eIdle;    // 相位待机 / phase idle
    _fTrimHeld   := 0.0;                       // 修正量保持量 0 [%] / held trim zero
    _bConfirmBreak := TRUE;                    // 节拍计时从零开始 / cadence timer starts from zero
    _bInit       := TRUE;                      // 首扫只做一次 / the first scan runs once
END_IF

(*------------------------------------------------------------------------------
 * 段 3｜参数闸门（四参数与冻结门限，任一非法即故障级；先于所有除法与比较）
 *      Parameter gate, any illegal value is a fault, checked before any arithmetic
 *-----------------------------------------------------------------------------*)
IF (fO2Target <> fO2Target) OR (ABS(fO2Target) > DL_VAL_LIM) OR (fO2Target <= DL_TARGET_MN) THEN
    _bParamBad := TRUE;                        // 目标氧含量非法 / target oxygen illegal
END_IF
IF (fO2Deadband <> fO2Deadband) OR (ABS(fO2Deadband) > DL_VAL_LIM) OR (fO2Deadband < DL_BAND_MN) THEN
    _bParamBad := TRUE;                        // 死区半宽非法 / dead band illegal
END_IF
IF (fTrimLimit <> fTrimLimit) OR (ABS(fTrimLimit) > DL_VAL_LIM) OR (fTrimLimit <= DL_LIMIT_MN) THEN
    _bParamBad := TRUE;                        // 修正限幅非法 / trim limit illegal
END_IF
IF (fTrimStep <> fTrimStep) OR (ABS(fTrimStep) > DL_VAL_LIM) OR (fTrimStep <= DL_STEP_MN) THEN
    _bParamBad := TRUE;                        // 步长非法 / step illegal
END_IF
IF (fRateFreeze <> fRateFreeze) OR (ABS(fRateFreeze) > DL_VAL_LIM) OR (fRateFreeze <= DL_RATE_MN) THEN
    _bParamBad := TRUE;                        // 冻结门限非法 / freeze threshold illegal
END_IF

(*------------------------------------------------------------------------------
 * 段 4｜输入有限性与偏差计算（区间判据同时拦 NaN 与 ±Inf）
 *      Input finiteness and deviation, the interval test catches NaN and infinity
 *-----------------------------------------------------------------------------*)
_fDev     := 0.0;                              // 偏差预置 0 [%] / deviation preset to zero
_fAbsDev  := 0.0;                              // 偏差绝对值预置 0 [%] / absolute deviation preset to zero
_fAbsRate := 0.0;                             // 负荷率绝对值预置 0 [%/s] / absolute load rate preset to zero

IF (fO2Meas < -DL_VAL_LIM) OR (fO2Meas > DL_VAL_LIM) THEN
    _bFiniteBad := TRUE;                       // 氧量非有限 / oxygen non-finite
END_IF
IF (fLoadRate < -DL_VAL_LIM) OR (fLoadRate > DL_VAL_LIM) THEN
    _bFiniteBad := TRUE;                       // 负荷率非有限 / load rate non-finite
END_IF

IF NOT _bFiniteBad THEN
    _fDev     := fO2Meas - fO2Target;           // 偏差：正 = 空气偏多 [%] / positive means too much air
    _fAbsDev  := ABS(_fDev);                    // 偏差绝对值 [%] / absolute deviation
    _fAbsRate := ABS(fLoadRate);                // 负荷率绝对值 [%/s] / absolute load rate
END_IF
_fBandUse := LIMIT(DL_BAND_MN, fO2Deadband, DL_O2_MAX); // 生效死区半宽钳进物理域 [%] / effective dead band clamped

(*------------------------------------------------------------------------------
 * 段 5｜定时器无条件刷新（R40：在 CASE 之外每拍必调；步进后断输入一拍重启节拍）
 *      Timer refreshed unconditionally outside the CASE, restarted after each step
 *-----------------------------------------------------------------------------*)
_tConfirmUse := tConfirm;                      // 确认时间直取引脚 [ms] / confirm time taken from the pin
IF TIME_TO_DINT(_tConfirmUse) > DL_CONF_MAX_MS THEN
    _tConfirmUse := DINT_TO_TIME(DL_CONF_MAX_MS); // 超上限钳位，无专用码位（R90 不新开码） / clamped, no dedicated code
END_IF
IF TIME_TO_DINT(_tConfirmUse) < 0 THEN
    _tConfirmUse := DL_TIME_ZERO;              // 负数时间结构性不可达，兜底为 0 / structurally unreachable, fallback to zero
END_IF

_bCond := bEnable AND (NOT _bParamBad) AND (NOT _bFiniteBad)
          AND (_fAbsDev > _fBandUse) AND (_fAbsRate <= fRateFreeze); // 步进条件 / step condition

fbConfirm(IN := _bCond AND (NOT _bConfirmBreak), PT := _tConfirmUse); // 节拍计时无条件刷新
_bConfirmBreak := FALSE;                       // 断输入拍在调用后自清（R40 自清位置） / break self-cleared after the call

IF _bCond AND (fbConfirm.Q OR (_tConfirmUse <= DL_TIME_ZERO)) THEN
    _bStepPulse := TRUE;                       // 本拍走一步（tConfirm = 0 时每拍一步，合法语义） / one step this scan
END_IF

(*------------------------------------------------------------------------------
 * 段 6｜相位机（只做迁移；修正量在段 7 单点演进）
 *      Phase machine, transitions only, the trim evolves in segment seven
 *-----------------------------------------------------------------------------*)
CASE _eState OF

    E_DL_O2TrimState.eIdle:                    // 待机：参数合法、输入有限且使能即进入
        IF _bParamBad OR _bFiniteBad THEN
            _eState := E_DL_O2TrimState.eFault; // 原因未消失，转故障 / the cause persists
        ELSIF bEnable THEN
            IF _fAbsRate > fRateFreeze THEN
                _eState := E_DL_O2TrimState.eFrozen; // 负荷剧变，直接进冻结 / load jumping, freeze directly
            ELSE
                _eState := E_DL_O2TrimState.eActive; // 进生效相 / enter the active phase
            END_IF
        END_IF

    E_DL_O2TrimState.eActive:                  // 生效：越死区才步进
        IF NOT bEnable THEN
            _eState := E_DL_O2TrimState.eIdle; // 失能回待机 / disabled, back to idle
        ELSIF _bParamBad OR _bFiniteBad THEN
            _eState := E_DL_O2TrimState.eFault; // 转故障 / go to fault
        ELSIF _fAbsRate > fRateFreeze THEN
            _eState := E_DL_O2TrimState.eFrozen; // 负荷剧变，冻结修正 / load jumping, freeze the trim
        END_IF

    E_DL_O2TrimState.eFrozen:                  // 冻结：负荷平稳后恢复
        IF NOT bEnable THEN
            _eState := E_DL_O2TrimState.eIdle; // 失能回待机 / disabled, back to idle
        ELSIF _bParamBad OR _bFiniteBad THEN
            _eState := E_DL_O2TrimState.eFault; // 转故障 / go to fault
        ELSIF _fAbsRate <= fRateFreeze THEN
            _eState := E_DL_O2TrimState.eActive; // 负荷已平稳，恢复修正 / load steady again, resume
        END_IF

    E_DL_O2TrimState.eFault:                   // 故障：原因消失即自动恢复（本件无复位引脚）
        IF NOT bEnable THEN
            _eState := E_DL_O2TrimState.eIdle; // 失能回待机 / disabled, back to idle
        ELSIF (NOT _bParamBad) AND (NOT _bFiniteBad) THEN
            IF _fAbsRate > fRateFreeze THEN
                _eState := E_DL_O2TrimState.eFrozen; // 原因消失但负荷仍剧变，进冻结 / cause cleared but the load still jumps
            ELSE
                _eState := E_DL_O2TrimState.eActive; // 原因消失自动回生效相 / cause cleared, resume
            END_IF
        END_IF

    ELSE
        _bIllegal := TRUE;                     // 标记非法状态 / flag the illegal state
        _eState   := E_DL_O2TrimState.eFault;  // 回故障态 / back to the fault state
END_CASE

(*------------------------------------------------------------------------------
 * 段 7｜修正量演进（仅生效相且本拍有步进脉冲；累加后双侧钳，钳位后不再累加）
 *      Trim evolution in the active phase only, clamped both ways right after the step
 *-----------------------------------------------------------------------------*)
IF (_eState = E_DL_O2TrimState.eActive) AND _bStepPulse THEN
    IF _fDev > _fBandUse THEN
        _fTrimHeld := _fTrimHeld - fTrimStep;  // 氧量偏高：减空气 [%] / oxygen high, reduce air
    ELSIF (_fBandUse - _fDev) > DL_EPS THEN
        _fTrimHeld := _fTrimHeld + fTrimStep;  // 氧量偏低：增空气 [%] / oxygen low, add air
    END_IF
    _fTrimHeld := LIMIT(-fTrimLimit, _fTrimHeld, fTrimLimit); // 抗饱和：双侧钳位，不回算积分 / anti-windup, clamp only
    _bConfirmBreak := TRUE;                    // 走一步后重启节拍，节拍严格等于 tConfirm / restart the cadence
END_IF

(*------------------------------------------------------------------------------
 * 段 8｜输出单点写入与码位优先级链
 *      Single write point of the outputs and the code priority chain
 *-----------------------------------------------------------------------------*)
IF _bIllegal THEN
    fTrim   := 0.0;                            // 非法状态：修正量归零 [%] / illegal state, trim zeroed
    bActive := FALSE;                          // 生效标志清零 / active flag cleared
    bFrozen := FALSE;                          // 冻结标志清零 / frozen flag cleared
    eErr    := 16#0002_2C12;                   // 故障级：状态机兜底 / fault: state machine fallback
    bError  := TRUE;                           // 置故障标志 / raise the fault flag
    bValid  := FALSE;                          // 输出不可用 / outputs unusable
ELSIF NOT bEnable THEN
    fTrim      := 0.0;                         // 失能：修正量显式清零 [%] / disabled, trim explicitly zeroed
    _fTrimHeld := 0.0;                         // 保持量一并清零，再使能不回投旧偏置 [%] / held trim cleared too
    bActive    := FALSE;                       // 生效标志清零 / active flag cleared
    bFrozen    := FALSE;                       // 冻结标志清零 / frozen flag cleared
    bValid     := FALSE;                       // 失能时输出不可用 / unusable while disabled
ELSIF _bParamBad THEN
    fTrim      := 0.0;                         // 参数非法：退回纯交叉限幅，修正量 0 [%] / trim zeroed, cross limiting only
    _fTrimHeld := 0.0;                         // 保持量清零，防非法参数解除后旧值回投 [%] / held trim cleared
    bActive    := FALSE;                       // 生效标志清零 / active flag cleared
    bFrozen    := FALSE;                       // 冻结标志清零 / frozen flag cleared
    eErr       := 16#0002_2C10;                // 故障级：修正参数非法 / fault: trim parameters illegal
    bError     := TRUE;                        // 置故障标志 / raise the fault flag
    bValid     := FALSE;                       // 输出不可用 / outputs unusable
ELSIF _bFiniteBad THEN
    fTrim   := _fTrimHeld;                     // 非有限：保持末次修正量 [%] / hold the last trim
    bActive := FALSE;                          // 本次未演进，不宣称生效 / no evolution this scan
    bFrozen := FALSE;                          // 本次未演进，不宣称冻结 / no freeze claim this scan
    eErr    := 16#0002_2C11;                   // 故障级：输入非有限 / fault: non-finite input
    bError  := TRUE;                           // 置故障标志 / raise the fault flag
    bValid  := FALSE;                          // 输出不可用 / outputs unusable
ELSE
    fTrim   := _fTrimHeld;                     // 正常：修正量出口 [%] / trim outlet
    bActive := (_eState = E_DL_O2TrimState.eActive); // 生效标志 / active flag
    bFrozen := (_eState = E_DL_O2TrimState.eFrozen); // 冻结标志 / frozen flag
    bValid  := TRUE;                           // 输出可用 / outputs usable
    IF _eState = E_DL_O2TrimState.eFrozen THEN
        eErr := 16#0002_2C02;                  // 信息级：负荷变化率超限已冻结 / informational: frozen by the load rate
    ELSIF _fAbsDev <= _fBandUse THEN
        eErr := 16#0002_2C01;                  // 信息级：死区内不修正 / informational: inside the dead band
    END_IF
END_IF

END_FUNCTION_BLOCK

(* ---- FB_DL_ExtremumSeekCtrl.st ---- *)
(*==============================================================================
 * 组件名称 (Component)  : FB_DL_ExtremumSeekCtrl
 * 所属子库 (Sublibrary) : DL_Algo
 * 当前版本 (Version)    : 1.0.1
 * 兼容性 (Platform)     : CODESYS 3.5+ / TwinCAT 3 / 汇川 InoProShop / 施耐德 Machine Expert
 *                         仅依赖 Standard.library（TON / SIN / ABS），零厂商私有库
 * 功能描述 (Function)   : 极值寻优控制（扰动观察式 ES，无需模型）。在设定点
 *                         上叠加正弦扰动 dith = fDithAmp·SIN(ω·t)，对输出量
 *                         y 做同步解调：梯度估计 g ≈ 均值(y·dith)/均方(dith²)
 *                         （滚动窗归一化互相关），g > 0 说明设定点应增大、
 *                         g < 0 应减小；积分器按 fStepGain·g 调整设定点，
 *                         fSetpointOut = fSetBase + fTrim。设定点漂移追踪、
 *                         燃烧效率寻优、光伏 MPPT 类场景（公开 ES 语义 clean-room）。
 * 来源标签 (Origin)     : 自研线（公开极值寻优算法语义 clean-room，IEC 61131-3
 *                         标准语义的道莅防御性实现，零代码行复制）
 * 边界语义 (Boundary)   : ① 归一化除零防御：窗内均方 dith² <= eps（扰动被禁
 *                         或窗未填充）→ 梯度按 0（设定点保持），不产生 Inf；
 *                         ② 输出 NaN/Inf 拒收：y 非有限拍不参与解调累计；
 *                         ③ 修剪限幅：fTrim 双侧钳位于 [-fTrimLimit, +fTrimLimit]
 *                         （R151 补偿量钳位口径），防梯度发散把设定点推飞；
 *                         ④ 组态闸：扰动幅值/增益/限幅域检查 → 故障锁存。
 * 输出语义 (Fallback)   : 【R191】bEnable = FALSE → 修剪保持（设定点不跳变，
 *                         扰动冻结），bDitherOut = FALSE；eFault 相 → 修剪保持
 *                         末值 + bError = TRUE。
 * 码位     (Codes)      : 按 R297 范式零 16# 码位硬编码；错误出口 BOOL+ENUM(eCause)，
 *                         码位待主控收口统一派号。
 * 红线自检 (Redline)    : 7 项红线已自检：R1 零全局 ✓｜R2 零物理地址 ✓｜R3 纯 IEC ✓
 *                         R4 除零（均方 eps 闸）/NaN 拒收/修剪钳位/组态闸 ✓
 *                         R5 双语同行注释 ✓｜R6 CASE 带 ELSE 兜底迁 eFault ✓
 *                         R7 TON/R_TRIG 段 0 无条件刷新 ✓
 * 验收向量 (Acceptance) : V1 y = -(x-50)² + 100（峰在 50），从 x=40 起寻优
 *                         → fTrim 单调逼近 +10（容差由 fStepGain/窗深决定）；
 *                         V2 峰左侧（g>0）→ fTrim 递增；峰右侧（g<0）→ 递减；
 *                         V3 fTrim 到 ±fTrimLimit 饱和不再外推。
 * 修订历史 (Revision)   : 2026-11-20  v1.0.0  R49 首版（批 3 · 序号 12）
 *                        2026-11-20  v1.0.1  R51 返修（R50 终审中×2）：①相位推进
 *                        删多乘 2.0 因子（扰动频率与组态周期一致）；②解调窗改真
 *                        滚动窗口径：tonWin 自复位（IN 带 NOT tonWin.Q，FB33-2），
 *                        到时单拍清 Σy·dith / Σdith² / 样本数，eIdle 相同步清窗，
 *                        梯度只反映最近 tWinTime 窗（与功能描述「滚动窗」一致）
 *==============================================================================*)
TYPE E_DL_EscState :
(
    eIdle  := 0,                             (* 待使能（修剪保持零） / Idle, trim held *)
    eSeek  := 10,                            (* 扰动寻优运行 / Perturb-and-seek run *)
    eFault := 90                             (* 故障锁存相 / Fault latched phase *)
);
END_TYPE

TYPE E_DL_EscCause :
(
    eNone       := 0,                        (* 无故障成因 / No cause *)
    eCfgIllegal := 1,                        (* 组态非法：扰动/增益/限幅越域 / Illegal config *)
    ePhaseBad   := 2                         (* 非法相位兜底 / Illegal phase fallback *)
);
END_TYPE

FUNCTION_BLOCK FB_DL_ExtremumSeekCtrl
VAR_INPUT
    fY          : LREAL := 0.0;              (* 寻优输出量（被最大化目标）[工程单位] / Objective output to maximize *)
    fDithAmp    : LREAL := 1.0;              (* 正弦扰动幅值，域 > 0.0 [工程单位] / Dither amplitude *)
    fDithPeriod : TIME := T#2S;              (* 扰动周期，域 >= 20·tScan 工程约束（组态闸按非零检查）[ms] / Dither period *)
    tWinTime    : TIME := T#5S;              (* 解调滚动窗保持时长，域 > T#0S [ms] / Demodulation window hold time *)
    fStepGain   : LREAL := 0.5;              (* 梯度→修剪积分增益，域 > 0.0 [工程单位/拍] / Step gain *)
    fTrimLimit  : LREAL := 10.0;             (* 修剪限幅，域 > 0.0 [工程单位] / Trim limit *)
    fScanS      : LREAL := 0.01;             (* 扫描周期秒值（相位推进步长），域 > 1E-6 [s] / Scan period seconds *)
    bEnable     : BOOL := TRUE;              (* 寻优使能，FALSE 修剪保持扰动冻结 [-] / Enable *)
    bReset      : BOOL := FALSE;             (* 复位命令，上升沿清修剪/窗/相位 [-] / Reset command *)
END_VAR
VAR_OUTPUT
    fSetpointOut : LREAL;                    (* 设定点输出 = 基准 + 修剪 [工程单位] / Setpoint output *)
    fDitherOut   : LREAL;                    (* 当前扰动瞬时值（注入量诊断镜像）[工程单位] / Dither instantaneous value *)
    fTrim        : LREAL;                    (* 当前修剪量（相对基准偏移）[工程单位] / Current trim *)
    fGradEst     : LREAL;                    (* 当前梯度估计（归一化互相关）[-] / Gradient estimate *)
    bWindowFull  : BOOL;                     (* 窗到时清窗单拍脉冲（滚动窗节拍指示）[-] / Window-expiry single-scan pulse *)
    eState       : E_DL_EscState;            (* 状态出口 / State outlet *)
    eCause       : E_DL_EscCause;            (* 故障成因出口（R190 归因唯一） / Fault cause outlet *)
    bError       : BOOL;                     (* 故障锁存标志 [-] / Fault latch flag *)
END_VAR
VAR
    _eState : E_DL_EscState := E_DL_EscState.eIdle;       (* 内部相位（CASE 唯一写入目标） / Internal phase *)
    _eCause : E_DL_EscCause := E_DL_EscCause.eNone;       (* 故障成因锁存量 / Latched cause *)
    rtReset : R_TRIG;                        (* 复位沿实例，段 0 无条件调用 / Reset edge instance *)
    tonWin  : TON;                           (* 解调窗计时，段 0 无条件调用 / Demod window timer *)
    _fPhase : LREAL := 0.0;                  (* 扰动相位累计（弧度），2π 回卷 [rad] / Dither phase accumulator *)
    _fDith  : LREAL;                         (* 本拍扰动瞬时值 [工程单位] / Dither this scan *)
    _fSxy   : LREAL;                         (* 解调窗累计：Σ y·dith [工程单位²] / Demod sum y·dith *)
    _fSdd   : LREAL;                         (* 解调窗累计：Σ dith² [工程单位²] / Demod sum dith² *)
    _nFill  : UDINT;                         (* 窗内有效样本数 [拍] / Valid sample count *)
    _fG     : LREAL;                         (* 本拍梯度估计 [-] / Gradient this scan *)
    _fTrimI : LREAL;                         (* 修剪量锁存（积分器）[工程单位] / Trim integrator latch *)
    _bFault : BOOL;                          (* 故障锁存位 / Latched fault bit *)
    _bCfgBad: BOOL;                          (* 组态非法当拍量 / Illegal config this scan *)
END_VAR
VAR CONSTANT
    DL_ESC_EPS    : LREAL := 1.0E-12;        (* 均方判零容差 [工程单位²] / Mean-square epsilon *)
    DL_ESC_2PI    : LREAL := 6.28318530717958648;   (* 2π（相位回卷界）[rad] / Two pi *)
    DL_ESC_TRIMMAX: LREAL := 1.0E6;          (* 修剪绝对安全上限（防积分器发散）[工程单位] / Trim absolute safety cap *)
    DL_ESC_NMAX   : UDINT := 4294960000;     (* 样本计数回绕防护上限 [-] / Sample count wrap guard *)
END_VAR

(* —— 段 0：当拍判据派生 + 实例无条件刷新（R228A） —— *)
_bCfgBad := (fDithAmp <= 0.0) OR (fStepGain <= 0.0) OR (fTrimLimit <= 0.0)   (* 组态闸：幅值/增益/限幅正域（R151 全引脚） / Config gate *)
            OR (fDithPeriod <= T#0S) OR (tWinTime <= T#0S) OR (fScanS <= 1.0E-6);
rtReset(CLK := bReset);                      (* 复位沿每拍必调 / Reset edge every scan *)
tonWin(IN := (_eState = E_DL_EscState.eSeek) AND NOT tonWin.Q, PT := tWinTime);   (* 解调滚动窗自复位计时（FB33-2：IN 带自身 Q 取反，到时单拍后自动重启） / Self-resetting window timer *)
IF tonWin.Q THEN                             (* 窗到时单拍：清解调累计（滚动窗口径，与头注释一致，R338） / Window expiry: clear demod sums *)
    _fSxy := 0.0;                            (* 清 Σy·dith / Clear demod sum *)
    _fSdd := 0.0;                            (* 清 Σdith² / Clear mean-square sum *)
    _nFill := 0;                             (* 清有效样本数 / Clear fill count *)
END_IF
_fPhase := _fPhase + DL_ESC_2PI * fScanS / (TIME_TO_LREAL(fDithPeriod) / 1000.0);   (* 相位推进：ω·dt（v1.0.1 删多乘 2.0 因子），除子为周期秒值（组态闸已保证 > 0），无除零 / Phase advance ω·dt, divisor gated *)
IF _fPhase >= DL_ESC_2PI THEN
    _fPhase := _fPhase - DL_ESC_2PI;         (* 相位 2π 回卷（防浮点精度坍缩） / Phase wrap *)
END_IF
_fDith := fDithAmp * SIN(_fPhase);           (* 本拍扰动值（标准 SIN） / Dither value *)

(* —— 段 1：单拍量预清零（R107） —— *)
_fG := 0.0;                                  (* 梯度缺省 0（未定语义：不驱动修剪） / Gradient default zero *)

(* —— 段 2：复位沿处理（作用域：清故障 + 清修剪积分器 + 清窗累计 + 清相位，R283 逐项声明） —— *)
IF rtReset.Q THEN
    _bFault := FALSE;                        (* 清故障锁存 / Clear fault *)
    _eCause := E_DL_EscCause.eNone;          (* 清成因 / Clear cause *)
    _fTrimI := 0.0;                          (* 清修剪积分器 / Clear trim integrator *)
    _fSxy := 0.0;                            (* 清解调累计 / Clear demod sums *)
    _fSdd := 0.0;                            (* 清均方累计 / Clear dith² sum *)
    _nFill := 0;                             (* 清样本数 / Clear fill count *)
    _fPhase := 0.0;                          (* 清相位 / Clear phase *)
    _eState := E_DL_EscState.eIdle;          (* 迁待机相 / Back to idle *)
END_IF

(* —— 段 3：组态闸故障锁存（R45 配对；锁存至复位沿，R189） —— *)
IF _bCfgBad AND NOT _bFault THEN
    _bFault := TRUE;                         (* 锁存故障位 / Latch fault *)
    _eCause := E_DL_EscCause.eCfgIllegal;    (* 成因：组态非法 / Cause: illegal config *)
    _eState := E_DL_EscState.eFault;         (* 同步迁故障相 / Migrate to fault *)
END_IF

(* —— 段 4：CASE 主状态机（ELSE 兜底迁 eFault，红线 6） —— *)
CASE _eState OF
    E_DL_EscState.eIdle:                     (* 待机相：修剪保持、扰动冻结 / Idle *)
        _fSxy := 0.0;                        (* 待机清窗：窗只含连续 eSeek 期样本（滚动窗口径） / Clear window while idle *)
        _fSdd := 0.0;                        (* 清 Σdith² / Clear mean-square sum *)
        _nFill := 0;                         (* 清有效样本数 / Clear fill count *)
        IF bEnable AND NOT _bFault THEN
            _eState := E_DL_EscState.eSeek;  (* 进入寻优 / Enter seek *)
        END_IF
    E_DL_EscState.eSeek:                     (* 寻优相：解调 + 梯度积分 / Seek *)
        IF NOT bEnable THEN
            _eState := E_DL_EscState.eIdle;  (* 失能回待机（修剪保持不回零） / Back to idle, trim held *)
        ELSE
            IF (fY = fY) AND ((fY - fY) = (fY - fY)) THEN   (* 输出有限（NaN 自反 + Inf 差判） / Finite objective *)
                _fSxy := _fSxy + fY * _fDith;   (* 解调累计 Σy·dith / Demod accumulate *)
                _fSdd := _fSdd + _fDith * _fDith;   (* 均方累计 Σdith² / Mean-square accumulate *)
                IF _nFill < DL_ESC_NMAX THEN
                    _nFill := _nFill + 1;    (* 有效样本计数（UDINT 回绕防护） / Sample count, wrap-guarded *)
                END_IF
            END_IF
            IF (_fSdd > DL_ESC_EPS) AND (_nFill >= 8) THEN   (* 归一化除零闸 + 最小样本闸（边界①） / Normalization gate *)
                _fG := _fSxy / _fSdd;        (* 梯度估计 = Σy·dith / Σdith²（同窗归一化互相关） / Gradient estimate *)
            END_IF
            _fTrimI := _fTrimI + fStepGain * _fG;   (* 梯度驱动修剪积分 / Gradient-driven trim integrate *)
            IF _fTrimI > fTrimLimit THEN
                _fTrimI := fTrimLimit;       (* 修剪上限钳位（R151 口径） / Trim upper clamp *)
            ELSIF _fTrimI < (-fTrimLimit) THEN
                _fTrimI := (-fTrimLimit);    (* 修剪下限钳位 / Trim lower clamp *)
            END_IF
            IF ABS(_fTrimI) > DL_ESC_TRIMMAX THEN
                _fTrimI := DL_ESC_TRIMMAX;   (* 绝对安全上限兜底（防组态限幅被绕过） / Absolute safety cap *)
            END_IF
        END_IF
    E_DL_EscState.eFault:                    (* 故障相：修剪与扰动冻结，仅复位沿出 / Fault *)
        ;                                    (* 锁存回放（R28） / Replay from latch *)
    ELSE                                     (* 非法相位兜底迁安全态 / Illegal phase fallback *)
        _eState := E_DL_EscState.eFault;     (* 迁故障相 / To fault *)
        _bFault := TRUE;                     (* 同步锁存 / Latch *)
        _eCause := E_DL_EscCause.ePhaseBad;  (* 成因：非法相位 / Cause: illegal phase *)
END_CASE

(* —— 段 5：出口映射（bError/eState 同源，R191） —— *)
fTrim := _fTrimI;                            (* 修剪出口镜像 / Trim mirror *)
fSetpointOut := _fTrimI;                     (* 设定点 = 修剪（基准由调用方叠加，属主边界：本件只管修剪量） / Setpoint = trim, base owned by caller *)
fDitherOut := _fDith;                        (* 扰动瞬时值镜像 / Dither mirror *)
fGradEst := _fG;                             (* 梯度估计镜像 / Gradient mirror *)
bWindowFull := tonWin.Q;                     (* 窗到时单拍脉冲镜像 / Window-expiry pulse mirror *)
bError := _bFault;                           (* 故障标志镜像 / Fault flag mirror *)
eState := _eState;                           (* 状态出口 / State outlet *)
eCause := _eCause;                           (* 成因出口 / Cause outlet *)
END_FUNCTION_BLOCK

(* ---- FB_DL_FanArraySeq.st ---- *)
// =====================================================================
// FB_DL_FanArraySeq.st
// 风机阵列轮值与变频/工频混拖调度（轮值均衡 + 分级投切 + 混拖互斥）
// Fan array duty rotation and VFD/direct staging scheduler
// 所属子库: DL_Algo    版本: v1.0.0    兼容: CODESYS V3.5+ / TwinCAT 3 / 汇川 InoProShop
// 码位: 16#0002_3729 ~ 16#0002_372D (本件独占 5 槽, 勿复用)
// 溯源: 道莅 clean-room 防御性实现
//       来源组标签: hvac, fan-array, duty-rotation, staging
// 修改记录: R30 初版 (ROUND_PLAN_R30 序 17)
// 分层声明: 本件为阵列级编排, 轮值均衡沿用库内轮值件范式、分级投切沿用
//           风机阵列分级件范式, 单台风机本体控制不在本件复现;
//           混拖互斥: 同一台风机同一拍至多处于变频或工频一种模式
// =====================================================================
FUNCTION_BLOCK FB_DL_FanArraySeq
VAR_INPUT
    bEnable    : BOOL  := FALSE;    // 使能 / Enable
    uReqStages : USINT := 2;        // 需求台数 0~6, 越界钳位 / Required stages, clamped
    abFanAvail : ARRAY[1..6] OF BOOL;   // 各台风机可用反馈 / Fan availability
    abVfdEn    : ARRAY[1..6] OF BOOL;   // 各台变频位（真 = 具备变频能力）/ VFD-capable flag
    tMinRun    : TIME  := T#30S;    // 最短运行时间（防振颤与轮值门槛）T#1S~T#60M / Min run time [s]
    bRotateReq : BOOL  := FALSE;    // 轮值请求命令 / Rotation request
END_VAR
VAR_OUTPUT
    abFanRun     : ARRAY[1..6] OF BOOL;   // 各台运行输出 / Fan run outputs
    abFanVfdMode : ARRAY[1..6] OF BOOL;   // 各台变频模式输出 / Fan VFD mode outputs
    uRunCount    : USINT := 0;      // 运行台数 / Running count
    eErr         : UDINT := 16#0002_3729;  // 错误码 / Error code
END_VAR
VAR
    rtrRotate  : R_TRIG;            // 轮值请求沿, 每拍无条件刷新 / Rotate edge, refreshed every cycle
    aTonRun    : ARRAY[1..6] OF TON;    // 各台运行计时, 每拍无条件刷新 / Per-fan run timers, refreshed every cycle
    abRunSel   : ARRAY[1..6] OF BOOL;   // 本拍期望运行集 / Desired run set this cycle
    uLeadIdx   : USINT := 1;       // 轮值起始索引 / Rotation lead index
    uReq       : USINT := 0;       // 钳位后需求台数 / Clamped demand
    uTarget    : USINT := 0;       // 实际目标台数 / Effective target
    uAvailCnt  : USINT := 0;       // 可用台数 / Available count
    uSelCnt    : USINT := 0;       // 已选台数 / Selected count
    uK         : USINT := 0;       // 轮转探测偏移 / Rotation probe offset
    uIdx       : USINT := 1;       // 轮转探测索引 / Rotation probe index
    uNext      : USINT := 1;       // 轮值推进探测索引 / Lead advance probe index
    uProbe     : USINT := 0;       // 轮值推进守卫计数 / Lead advance guard counter
    bClamp     : BOOL := FALSE;     // 需求越界钳位标记 / Demand clamp flag
    bShort     : BOOL := FALSE;     // 需求超可用标记 / Demand exceeds availability flag
    bRotOk     : BOOL := FALSE;     // 轮值允许标记 / Rotation allowed flag
    bStarted   : BOOL := FALSE;     // 本拍已投一台标记 / Started one this cycle flag
    bStopped   : BOOL := FALSE;     // 本拍已停一台标记 / Stopped one this cycle flag
    uZi        : INT   := 1;       // 1..6 数组下标 / Array subscript 1..6
END_VAR

// ---------------------------------------------------------------------
// 代码位表（本件独占, 勿复用）:
//   16#0002_3729 信息 阵列调度正常
//   16#0002_372A 信息 需求台数越界钳位（大于 6 已钳到 6）
//   16#0002_372B 信息 需求超可用（只投可用台数, 缺口提示）
//   16#0002_372C 信息 轮值等待（存在未达最短运行时间的运行台, 轮值请求挂起）
//   16#0002_372D 信息 待机未使能（全停安全侧）
// ---------------------------------------------------------------------

// ---- 需求钳位 / Demand clamp ----
bClamp := FALSE;
uReq := uReqStages;
IF uReqStages > 6 THEN
    uReq := 6;                      // 上界钳位 / Clamp upper
    bClamp := TRUE;                 // 置钳位信息 / Set clamp info
END_IF

// ---- 可用台数 / Available count ----
uAvailCnt := 0;
FOR uZi := 1 TO 6 DO
    IF abFanAvail[uZi] THEN
        uAvailCnt := uAvailCnt + 1;
    END_IF
END_FOR

// ---- 目标台数（不超可用, 台数 0 → 全停安全侧）/ Effective target ----
uTarget := uReq;
IF uTarget > uAvailCnt THEN
    uTarget := uAvailCnt;           // 只投可用数 / Only available count
    bShort := TRUE;                 // 置缺口信息 / Set shortfall info
END_IF

// ---- 轮值沿与运行计时实例无条件周期刷新 / Unconditional edge and timer refresh ----
rtrRotate(CLK := bRotateReq);
FOR uZi := 1 TO 6 DO
    aTonRun[uZi](IN := abFanRun[uZi], PT := tMinRun);   // 运行计时 / Run timing
END_FOR

// ---- 未使能全停（安全侧）/ All stop when disabled ----
IF NOT bEnable THEN
    FOR uZi := 1 TO 6 DO
        abFanRun[uZi] := FALSE;     // 全停 / All stop
    END_FOR
END_IF

// ---- 轮值允许判: 全部运行台已达最短运行时间 / Rotation allowed judge ----
bRotOk := TRUE;
FOR uZi := 1 TO 6 DO
    IF abFanRun[uZi] AND (NOT aTonRun[uZi].Q) THEN
        bRotOk := FALSE;            // 存在未达门槛的运行台 / Some fan below min run
    END_IF
END_FOR

// ---- 轮值推进: 全部运行台达门槛时沿探测推进起始索引（守卫计数防死循环）
//      Lead advance on rotation request ----
IF rtrRotate.Q AND bEnable AND bRotOk THEN
    uNext := uLeadIdx;              // 自当前起始索引探测 / Probe from lead
    uProbe := 0;
    WHILE uProbe < 6 DO
        uNext := uNext + 1;
        IF uNext > 6 THEN
            uNext := 1;             // 回绕 / Wrap
        END_IF
        uProbe := uProbe + 1;
        IF abFanAvail[uNext] THEN
            uLeadIdx := uNext;      // 推进起始索引 / Advance lead
            uProbe := 6;            // 提前退出 / Early exit
        END_IF
    END_WHILE
END_IF

// ---- 分级投切选择: 变频台优先, 轮值序探测, 工频补位 / Staging selection ----
FOR uZi := 1 TO 6 DO
    abRunSel[uZi] := FALSE;         // 期望集清空 / Clear desired set
END_FOR
uSelCnt := 0;
IF bEnable AND (uTarget > 0) THEN
    // 第一遍: 沿轮值序选变频台 / Pass 1: VFD-capable fans in rotation order
    uK := 0;
    WHILE (uK < 6) AND (uSelCnt < uTarget) DO
        uIdx := uLeadIdx + uK;
        IF uIdx > 6 THEN
            uIdx := uIdx - 6;       // 条件回绕, 不用取余 / Conditional wrap
        END_IF
        uK := uK + 1;
        IF abFanAvail[uIdx] AND abVfdEn[uIdx] AND (NOT abRunSel[uIdx]) THEN
            abRunSel[uIdx] := TRUE;
            uSelCnt := uSelCnt + 1;
        END_IF
    END_WHILE
    // 第二遍: 沿轮值序用工频台补位 / Pass 2: direct-on-line fans fill
    uK := 0;
    WHILE (uK < 6) AND (uSelCnt < uTarget) DO
        uIdx := uLeadIdx + uK;
        IF uIdx > 6 THEN
            uIdx := uIdx - 6;
        END_IF
        uK := uK + 1;
        IF abFanAvail[uIdx] AND (NOT abRunSel[uIdx]) THEN
            abRunSel[uIdx] := TRUE;
            uSelCnt := uSelCnt + 1;
        END_IF
    END_WHILE
END_IF

// ---- 分级投切执行: 同拍至多投一台、停一台（防振颤, 未达门槛不停机）
//      Staged apply: at most one start and one stop per cycle ----
bStarted := FALSE;
bStopped := FALSE;
FOR uZi := 1 TO 6 DO
    IF abRunSel[uZi] AND (NOT abFanRun[uZi]) AND (NOT bStarted) THEN
        abFanRun[uZi] := TRUE;      // 投入一台 / Start one
        bStarted := TRUE;
    END_IF
END_FOR
FOR uZi := 1 TO 6 DO
    IF (NOT abRunSel[uZi]) AND abFanRun[uZi] AND aTonRun[uZi].Q AND (NOT bStopped) THEN
        abFanRun[uZi] := FALSE;     // 停运一台（已达最短运行时间才停）/ Stop one eligible
        bStopped := TRUE;
    END_IF
END_FOR

// ---- 混拖模式输出（一台一拍至多一种模式）/ Mode outputs, one mode per fan ----
FOR uZi := 1 TO 6 DO
    abFanVfdMode[uZi] := abFanRun[uZi] AND abVfdEn[uZi];
END_FOR

// ---- 运行台数 / Running count ----
uRunCount := 0;
FOR uZi := 1 TO 6 DO
    IF abFanRun[uZi] THEN
        uRunCount := uRunCount + 1;
    END_IF
END_FOR

// ---- 错误码仲裁 / Error arbitration ----
IF NOT bEnable THEN
    eErr := 16#0002_372D;           // 待机全停 / Standby all stop
ELSIF bClamp THEN
    eErr := 16#0002_372A;           // 需求钳位 / Demand clamped
ELSIF bShort THEN
    eErr := 16#0002_372B;           // 需求超可用 / Short of availability
ELSIF bRotateReq AND (NOT bRotOk) THEN
    eErr := 16#0002_372C;           // 轮值等待 / Rotation pending
ELSE
    eErr := 16#0002_3729;           // 调度正常 / Normal
END_IF

END_FUNCTION_BLOCK

(* ---- FB_DL_FanPressureTrim.st ---- *)
(*
  FB_DL_FanPressureTrim  —  风机静压微调（偏差积分微调 + 抗饱和回退） / Fan static-pressure trim with integral adjustment and anti-windup back-off
  分类 Category : DL_Algo
  版本 Version  : 1.0.0
  来源 Source   : t2-7-packml — 包装线风系统微调算法深化
  溯源 Origin   : 道莅 clean-room 实现；死区 + 积分微调 + 饱和回退（条件积分抗饱和）为公开过程控制算法，未复制任何源码行
  功能 Function : 1) 偏差 _fErrKpa = fSpKpa - fPvKpa；2) 死区内（|偏差| <= fDeadbandKpa）冻结积分；
                  3) 积分微调：_fIntKpa += fKiKpaPerS × Δt（Δt 由 tCycle 换算，除数 1000.0 常量）；
                  4) 输出 = fTrimBaseKpa + _fIntKpa，钳制 [fOutMinKpa, fOutMaxKpa]；
                  5) 抗饱和回退：输出已顶上限且偏差仍为正（同向推高）时回退本周期积分增量；
                  输出已抵下限且偏差仍为负时同样回退，禁止积分继续累积（条件积分法）；
                  6) 上拍积分快照 _fIntPrevKpa 保存（R19 累计量快照，禁跨拍重算）；
                  7) 本件只有故障码、无信息码（派单硬约束）。
  接口 Interface: 输入设定/反馈/基准/增益/死区/周期/上下限；输出微调输出与积分镜像
  边界 Boundary : ① 组态闸：tCycle <= T#0S、fKiKpaPerS < 0.0、fDeadbandKpa < 0.0、
                  fOutMaxKpa <= fOutMinKpa → 038A 锁存；
                  ② 设定或反馈非有限（NaN 自反 + Inf 差值自减）→ 038A 锁存，输出冻结保持上一值
                  （R191：冻结保持，不降级置标志）；
                  ③ 积分器本身为限幅量，回退后仍钳制在 [fIntMinKpa, fIntMaxKpa] 域内；
                  ④ 浮点判据全容差式；⑤ 仅一个 R_TRIG 复位沿，段 0 无条件调用；
                  ⑥ 故障相迁出唯一路径 = bReset 上升沿；⑦ 零全局耦合（无 GVL / %I %Q %M）。
  依赖 Depends  : Standard.library（R_TRIG）
  码表 Error codes（Algo 段 0002，故障窗口 038A；本件无信息码）:
    16#0002_038A 故障级：静压微调故障总码（组态非法 / 设定或反馈非有限），
                 锁存至 bReset 上升沿；归因见 eCause，不新增码位（派单硬约束单码）
  修订历史 Revision :
    2026-11-19  v1.0.0  R43 首版（批次 3 · 序号 14）
*)

TYPE E_DL_FptState :
(
    eIdle  := 0,      // 未使能：输出冻结 / Idle, output frozen
    eRun   := 10,     // 微调运行中 / Trim active
    eFault := 90      // 故障锁存相（输出冻结保持） / Fault latched, output frozen
);
END_TYPE

TYPE E_DL_FptCause :
(
    eNone       := 0, // 无故障成因 / No cause
    eCfgIllegal := 1, // 组态非法 / Illegal configuration
    eNonFinite  := 2  // 设定或反馈非有限 / Non-finite setpoint or feedback
);
END_TYPE

FUNCTION_BLOCK FB_DL_FanPressureTrim
VAR_INPUT
    fSpKpa       : REAL := 0.0;        // 静压设定 [kPa] / Static pressure setpoint
    fPvKpa       : REAL := 0.0;        // 静压反馈 [kPa] / Static pressure feedback
    fTrimBaseKpa : REAL := 200.0;      // 微调基准输出 [kPa] / Trim base output
    fKiKpaPerS   : REAL := 0.5;        // 积分增益 [kPa/s]，域 >= 0 / Integral gain
    fDeadbandKpa : REAL := 2.0;        // 偏差死区 [kPa]，域 >= 0 / Deviation deadband
    fIntMinKpa   : REAL := -50.0;      // 积分量下限 [kPa] / Integral low limit
    fIntMaxKpa   : REAL := 50.0;       // 积分量上限 [kPa] / Integral high limit
    fOutMinKpa   : REAL := 100.0;      // 输出下限 [kPa] / Output low limit
    fOutMaxKpa   : REAL := 400.0;      // 输出上限 [kPa] / Output high limit
    tCycle       : TIME := T#100MS;    // 调用周期 [ms]，域 > 0 / Task cycle
    bEnable      : BOOL := FALSE;      // 微调使能（电平）[-] / Trim enable
    bReset       : BOOL := FALSE;      // 复位命令，上升沿清故障 [-] / Reset edge
END_VAR
VAR_OUTPUT
    eState       : E_DL_FptState;      // 状态出口，段 6 单点映射 / State outlet
    eCause       : E_DL_FptCause;      // 故障成因出口（R190） / Fault cause outlet
    fOutKpa      : REAL;               // 微调输出 [kPa] / Trim output
    fIntKpa      : REAL;               // 积分量镜像 [kPa] / Integral mirror
    bWindup      : BOOL;               // 抗饱和回退生效镜像 [-] / Anti-windup back-off mirror
    bError       : BOOL;               // 故障锁存标志 [-] / Fault latch flag
    nErrId       : UDINT;              // 故障码，0 = 无故障（本件无信息码） / Fault code only
END_VAR
VAR
    _eState      : E_DL_FptState := E_DL_FptState.eIdle;   // 内部相位（CASE 唯一写入目标） / Internal phase
    _eCause      : E_DL_FptCause := E_DL_FptCause.eNone;   // 故障成因锁存（锁存量） / Latched cause
    rtReset      : R_TRIG;             // 复位沿实例，每周期无条件调用 / Reset edge
    _fIntKpa     : REAL;               // 积分器保持量（持久） / Integral holding slot
    _fIntPrevKpa : REAL;               // 上拍积分快照（R19 累计量快照） / Previous-scan integral snapshot
    _fOutKpa     : REAL;               // 输出保持量（持久） / Output holding slot
    _fErrKpa     : REAL;               // 偏差 [kPa]（当拍量） / Deviation
    _fDeltaKpa   : REAL;               // 本周期积分增量 [kPa]（当拍量） / Integral increment
    _fOutCandKpa : REAL;               // 未钳制候选输出 [kPa]（当拍量） / Unclamped candidate
    _bWindupOn   : BOOL;               // 抗饱和回退当拍量 [-] / Anti-windup flag
    _bNonFin     : BOOL;               // 输入非有限当拍量 [-] / Non-finite input
    _bCfgBad     : BOOL;               // 组态非法当拍量 [-] / Config illegal
    _bFault      : BOOL;               // 故障锁存位（锁存量） / Latched fault bit
    _uFault      : UDINT;              // 故障码锁存（锁存量） / Latched fault code
END_VAR

(* —— 段 0：沿实例无条件周期刷新 + 当拍量判据 —— *)
_fErrKpa := fSpKpa - fPvKpa;                                                // 偏差 [kPa] / Deviation
_bNonFin := (fSpKpa <> fSpKpa) OR (fPvKpa <> fPvKpa)
         OR ((fSpKpa - fSpKpa) <> (fSpKpa - fSpKpa))
         OR ((fPvKpa - fPvKpa) <> (fPvKpa - fPvKpa));                       // NaN 自反 + Inf 差值自减 / NaN and Inf
_bCfgBad := (tCycle <= T#0S) OR (fKiKpaPerS < 0.0) OR (fDeadbandKpa < 0.0)
            OR (fOutMaxKpa <= fOutMinKpa) OR (fIntMaxKpa <= fIntMinKpa);    // 组态非法当拍量 / Config illegal
rtReset(CLK := bReset);                                                     // 复位沿，每拍必调 / Reset edge
_fIntPrevKpa := _fIntKpa;                                                   // 上拍积分快照（每拍无条件） / Previous integral snapshot

(* —— 段 1：单拍量预清零（锁存量与积分/输出保持槽不入清单） —— *)
bWindup := FALSE;                  // 抗饱和镜像缺省 FALSE / Anti-windup default
nErrId := 16#0000_0000;            // 故障码缺省无故障 / Fault code default

(* —— 段 2：复位沿 + 组态域闸 —— *)
IF rtReset.Q THEN                              // rtReset.Q = 当拍量 / current scan
    _bFault := FALSE;                          // 清故障锁存位（锁存量） / Clear fault latch
    _uFault := 16#0000_0000;                   // 清故障锁存码（锁存量） / Clear fault code
    _eCause := E_DL_FptCause.eNone;            // 清成因（锁存量） / Clear cause
    _fIntKpa := 0.0;                           // 清积分器 / Clear integrator
    _fIntPrevKpa := 0.0;                       // 清积分快照 / Clear snapshot
    IF _eState = E_DL_FptState.eFault THEN
        _eState := E_DL_FptState.eIdle;        // 故障相迁出：回未使能 / Fault exit to idle
    END_IF
END_IF
IF _bCfgBad THEN                               // 组态域闸 / Config gate
    _uFault := 16#0002_038A;                   // 故障级：微调故障总码 / Algo fault code
    _eCause := E_DL_FptCause.eCfgIllegal;      // 归因：组态非法 / Cause: illegal config
    _bFault := TRUE;                           // 标志与码位配对（R45） / Flag paired with code
END_IF
IF (NOT _bFault) AND _bNonFin THEN             // 非有限锁存 / Non-finite latch
    _uFault := 16#0002_038A;
    _eCause := E_DL_FptCause.eNonFinite;       // 归因：非有限 / Cause: non-finite
    _bFault := TRUE;
END_IF

(* —— 段 3：积分微调 + 抗饱和回退 + 输出钳制（仅运行相且无故障） —— *)
IF (NOT _bFault) AND (_eState = E_DL_FptState.eRun) THEN
    IF ABS(_fErrKpa) <= fDeadbandKpa THEN                    // 死区内：冻结积分（不动作） / Deadband freezes integrator
        _fDeltaKpa := 0.0;
    ELSE
        _fDeltaKpa := fKiKpaPerS * (TIME_TO_REAL(tCycle) / 1000.0);   // 周期加权积分增量（除常量 1000.0） / Cycle-weighted increment
        IF _fErrKpa < 0.0 THEN                               // 偏差为负：积分反向 / Negative deviation subtracts
            _fDeltaKpa := -_fDeltaKpa;
        END_IF
        _fIntKpa := _fIntKpa + _fDeltaKpa;                   // 积分累加 / Integrate
        IF _fIntKpa < fIntMinKpa THEN                        // 积分下限钳制 / Integral low clamp
            _fIntKpa := fIntMinKpa;
        ELSIF _fIntKpa > fIntMaxKpa THEN                     // 积分上限钳制 / Integral high clamp
            _fIntKpa := fIntMaxKpa;
        END_IF
    END_IF
    _fOutCandKpa := fTrimBaseKpa + _fIntKpa;                 // 候选输出 / Candidate output
    IF _fOutCandKpa > fOutMaxKpa THEN                        // 顶上限 / Hit high limit
        IF _fErrKpa > 0.0 THEN                               // 偏差仍同向推高：回退本周期增量 / Same-direction saturation
            _fIntKpa := _fIntPrevKpa;                        // 抗饱和回退到上拍快照 / Back-off to snapshot
            _bWindupOn := TRUE;
        END_IF
        _fOutKpa := fOutMaxKpa;                              // 输出钳制上限 / Output clamped high
    ELSIF _fOutCandKpa < fOutMinKpa THEN                     // 抵下限 / Hit low limit
        IF _fErrKpa < 0.0 THEN                               // 偏差仍同向推低：回退 / Same-direction saturation
            _fIntKpa := _fIntPrevKpa;                        // 抗饱和回退 / Back-off
            _bWindupOn := TRUE;
        END_IF
        _fOutKpa := fOutMinKpa;                              // 输出钳制下限 / Output clamped low
    ELSE
        _fOutKpa := _fOutCandKpa;                            // 未饱和：直接跟随 / Follow candidate
    END_IF
END_IF

(* —— 段 4：故障解除式（R240；全当拍量）：rtReset.Q / NOT _bCfgBad / NOT _bNonFin —— *)
IF rtReset.Q AND (NOT _bCfgBad) AND (NOT _bNonFin) THEN
    _bFault := FALSE;                          // 清故障锁存位（锁存量） / Clear fault latch
    _uFault := 16#0000_0000;                   // 清故障锁存码（锁存量） / Clear fault code
    _eCause := E_DL_FptCause.eNone;            // 清成因（锁存量） / Clear cause
END_IF

(* —— 段 4A：故障锁存相位迁移闸（输出冻结保持上一值） —— *)
IF _bFault AND (_eState <> E_DL_FptState.eFault) THEN
    _eState := E_DL_FptState.eFault;           // 锁存即入故障相 / Latch enters fault phase
END_IF

(* —— 段 5：相位机（CASE 全覆盖 + ELSE 兜底） —— *)
CASE _eState OF

E_DL_FptState.eIdle:
    IF bEnable AND (NOT _bFault) THEN          // 使能条件 / Enable gate
        _fIntKpa := 0.0;                       // 起始清积分（无扰切换） / Reset integrator on start
        _fOutKpa := fTrimBaseKpa;              // 起始输出取基准并钳制 / Start from base
        IF _fOutKpa < fOutMinKpa THEN
            _fOutKpa := fOutMinKpa;
        ELSIF _fOutKpa > fOutMaxKpa THEN
            _fOutKpa := fOutMaxKpa;
        END_IF
        _eState := E_DL_FptState.eRun;         // 进运行相 / Enter run
    END_IF

E_DL_FptState.eRun:
    IF NOT bEnable THEN                        // 撤使能：输出冻结，回未使能 / Disable: freeze and idle
        _eState := E_DL_FptState.eIdle;
    END_IF

E_DL_FptState.eFault:
    ;                                          // 故障相：输出冻结保持，仅段 4 复位沿可迁出 / Frozen, reset only

ELSE
    _uFault := 16#0002_038A;                   // 故障级：非法相位兜底（归并总码） / Illegal phase fallback
    _eCause := E_DL_FptCause.eCfgIllegal;      // 归因：相位非法归并组态 / Cause: phase illegal
    _bFault := TRUE;
    _eState := E_DL_FptState.eFault;           // 强制回故障相 / Force fault phase

END_CASE

(* —— 段 6：出口单点映射（名实同源；锁存码回放） —— *)
fOutKpa := _fOutKpa;                           // 输出出口 / Output outlet
fIntKpa := _fIntKpa;                           // 积分镜像 / Integral mirror
IF _bFault THEN
    nErrId := _uFault;                         // 故障锁存码回放 / Replay latched code
    bWindup := FALSE;                          // 故障相抗饱和镜像强制 FALSE / Anti-windup forced false
ELSE
    nErrId := 16#0000_0000;                    // 无故障：本件无信息码 / No fault, no info code
    bWindup := _bWindupOn;                     // 抗饱和镜像 / Anti-windup mirror
END_IF
bError := _bFault;                             // 故障标志同源 / Flag from latch
eState := _eState;                             // 状态出口 / State outlet
eCause := _eCause;                             // 成因出口 / Cause outlet

END_FUNCTION_BLOCK

(* ---- FB_DL_FanSurgeMarginCalc.st ---- *)
//==============================================================================
// 功能块：FB_DL_FanSurgeMarginCalc ｜ 中文名称：风机喘振裕度在线计算与分级预警
// 所属子库：DL_Algo ｜ 版本：v1.0.0 ｜ 日期：2026-11-23
// 兼容：CODESYS V3.5+ / TwinCAT 3 / 汇川 InoProShop（纯 IEC 61131-3 第 3 版，零方言）
// 功能描述：以线性化喘振线 p_surge(Q) = P0 − K·Q（零流量喘振压力 P0、斜率 K
//           引脚注入）在线计算风机工况点裕度：
//           fMarginPct = (p_surge − p_act)/p_surge × 100 [%]，
//           并按两级阈值分级：裕度 ≤ 预警阈 → eWarn（延时确认）；裕度 ≤ 跳机
//           阈或裕度 < 0（工况点越线）→ eTrip（跳机保护，锁存需复位沿解除）。
//           预警/跳机均经 TON 去抖确认，防喘振开环余量监视用途；闭环防喘振
//           放空阀调节不属本件职责。
// 开源溯源 (Origin)：原创实现（风机性能曲线公开口径，自研线，零外部源码行，
//           clean-room 独立编写）
// 公开接口清单：输入 bEn / bReset / fFlowAct / fPressAct / fSurgeP0 / fSurgeK /
//               fWarnMargin / fTripMargin / tWarnDelay / tTripDelay；
//               输出 fMarginPct / eLevel / bWarn / bTrip / uErrCode / bError / bValid
// 错误码表：16#0002_3920 信息级（裕度进入预警带，不置 bError）/
//           16#0002_3921 故障级（喘振线参数非法：P0 <= 0、K < 0 或非有限，
//           置 bError）/
//           16#0002_3922 信息级（工况点输入非有限，保持现状不置 bError）/
//           16#0002_3923 预留禁用（不得挪用）
// 状态机：E_DL_SurgeLevel（本文件唯一定义，全库唯一属主）：
//           eNormal = 0 / eWarn = 1 / eTrip = 2；非法分级兜底归 eTrip（安全侧）
// 边界行为：① P0 <= 0 或 K < 0 → 故障 3921 + bError，裕度输出 0；
//           ② 工况点非有限 → 信息 3922，bValid := FALSE，分级冻结；
//           ③ p_surge(Q) <= 容差（深越线）→ 分母闸钳容差，裕度深度负值照算；
//           ④ bTrip 锁存至 bReset 上升沿或撤使能（R189：锁存码有可达清除沿）；
//           ⑤ TON ×2 / R_TRIG ×1 每拍无条件刷新（不入分支，红线 R7）；
//           ⑥ CASE 带 ELSE，非法值兜底归 eTrip（安全侧）。
// 修订历史：v1.0.0 2026-11-23 首版（R73 派单 · 批 1 · 序 3）
//==============================================================================

(*------------------------------------------------------------------------------
 * 枚举: E_DL_SurgeLevel（归属本功能块，同文件发布，全库唯一属主）
 * 含义: 喘振裕度分级，成员与 CASE 标签双向完备。
 *-----------------------------------------------------------------------------*)
TYPE E_DL_SurgeLevel :
(
    eNormal := 0,    // 正常：裕度高于预警阈 / Normal, margin above the warning threshold
    eWarn   := 1,    // 预警：裕度进入预警带（延时确认）/ Warning band, delay confirmed
    eTrip   := 2     // 跳机：裕度越过跳机阈或越线（锁存）/ Trip band or beyond the line, latched
);
END_TYPE

(*==============================================================================
 * 功能块: FB_DL_FanSurgeMarginCalc
 * 调用约定: 每个扫描周期无条件调用一次；实例状态全部驻留于私有变量。
 * 调用示例: surgeWatch(fFlowAct := fFTx, fPressAct := fPTx,
 *                      fSurgeP0 := 12000.0, fSurgeK := 8.0,
 *                      fWarnMargin := 10.0, fTripMargin := 5.0);
 *          bWarn 接声光预警，bTrip 接防喘振放空联锁（开环余量监视）。
 * 组装说明: ① 喘振线参数须由工艺专业给值后引脚注入，禁在调用侧写
 *             魔法数（本件常量区只存防御参数）；
 *           ② bTrip 为锁存量，复位须经操作员确认沿 bReset 或撤使能；
 *           ③ 工况点测量引脚经 PRG_IoMapping 读入注入，本件零物理地址。
 *==============================================================================*)
FUNCTION_BLOCK FB_DL_FanSurgeMarginCalc
VAR_INPUT
    bEn         : BOOL := FALSE;      // 使能（FALSE 解除锁存回正常）/ Enable, FALSE releases the latch
    bReset      : BOOL := FALSE;      // 跳机锁存复位输入（上升沿有效）/ Trip latch reset, rising edge active
    fFlowAct    : LREAL := 0.0;       // 实测流量 [m3/h]，工况点横轴 / Measured flow [m3/h], operating point abscissa
    fPressAct   : LREAL := 0.0;       // 实测出口压 [Pa]，工况点纵轴 / Measured outlet pressure [Pa], operating point ordinate
    fSurgeP0    : LREAL := 12000.0;   // 零流量喘振压力 [Pa]，喘振线截距 / Surge line intercept at zero flow [Pa]
    fSurgeK     : LREAL := 8.0;       // 喘振线斜率 [Pa/(m3/h)]，右降为正 / Surge line slope [Pa per m3/h], positive falling
    fWarnMargin : LREAL := 10.0;      // 预警阈值 [百分数] / Warning margin threshold [percent]
    fTripMargin : LREAL := 5.0;       // 跳机阈值 [百分数] / Trip margin threshold [percent]
    tWarnDelay  : TIME := T#500MS;    // 预警去抖确认延时 [ms] / Warning debounce delay [ms]
    tTripDelay  : TIME := T#200MS;    // 跳机去抖确认延时 [ms] / Trip debounce delay [ms]
END_VAR
VAR_OUTPUT
    fMarginPct  : LREAL;              // 喘振裕度 [百分数]，正值安全 / Surge margin [percent], positive is safe
    eLevel      : E_DL_SurgeLevel;    // 分级结论 / Level conclusion
    bWarn       : BOOL;               // 预警声明（延时确认后）/ Warning declared after debounce
    bTrip       : BOOL;               // 跳机声明（锁存至复位沿）/ Trip declared, latched until reset edge
    uErrCode    : UDINT;              // 错误码，0 = 无错 / Error code, 0 = no error
    bError      : BOOL;               // 故障级标志，仅故障级错误置位 / Fault-class flag, set only on fault-level codes
    bValid      : BOOL;               // 输出可用标志 / Outputs usable flag
END_VAR
VAR
    tonWarn     : TON;                // 预警去抖定时器，每拍无条件刷新 / Warning debounce timer, refreshed every scan
    tonTrip     : TON;                // 跳机去抖定时器，每拍无条件刷新 / Trip debounce timer, refreshed every scan
    trigReset   : R_TRIG;             // 复位沿检测，每拍无条件刷新 / Reset edge detector, refreshed every scan
    fPSurge     : LREAL;              // 当前流量下喘振线压力 [Pa] / Surge line pressure at current flow [Pa]
    bInWarnBand : BOOL;               // 本拍裕度处于预警带（未确认）/ Margin in the warning band this scan, unconfirmed
    bInTripBand : BOOL;               // 本拍裕度处于跳机带或越线（未确认）/ Margin in the trip band or beyond, unconfirmed
END_VAR
VAR CONSTANT
    DL_SG_EPS   : LREAL := 1.0E-9;    // 浮点容差与分母闸 [Pa] / Float tolerance and denominator gate [Pa]
    DL_SG_INF   : LREAL := 1.7976931348623157E308; // LREAL 幅值上限 / LREAL magnitude ceiling
    DL_SG_PCT100: LREAL := 100.0;     // 裕度百分比放大系数 [1] / Margin percentage scale [1]
END_VAR

// ---- 段 1｜定时/沿实例无条件刷新（红线 R7：禁入条件分支）----
tonWarn(IN := bInWarnBand AND NOT bTrip, PT := tWarnDelay);   // 预警去抖按未确认态断输入 / Warning timer input per unconfirmed band
tonTrip(IN := bInTripBand AND NOT bTrip, PT := tTripDelay);   // 跳机去抖按未确认态断输入 / Trip timer input per unconfirmed band
trigReset(CLK := bReset);             // 复位沿每拍刷新 / Reset edge refreshed every scan

// ---- 段 2｜出口默认值：入口即赋确定值 ----
fMarginPct := 0.0;                    // 裕度默认零 / Margin preset zero
bWarn      := FALSE;                  // 预警默认 FALSE / Warning preset FALSE
uErrCode   := 16#0000_0000;           // 错误码先清零（信息级每拍重算）/ Error code cleared, info level recomputed
bError     := FALSE;                  // 故障标志先清零（R45 配对）/ Fault flag cleared first, R45 pairing
bValid     := FALSE;                  // 可用标志先清零 / Usable flag cleared first
bInWarnBand := FALSE;                 // 预警带声明先清零 / Warning band flag cleared first
bInTripBand := FALSE;                 // 跳机带声明先清零 / Trip band flag cleared first

// ---- 段 3｜喘振线参数闸：非法 → 故障 3921（R45 配对置 bError）----
IF (fSurgeP0 <> fSurgeP0) OR (ABS(fSurgeP0) > DL_SG_INF)
   OR (fSurgeK <> fSurgeK) OR (ABS(fSurgeK) > DL_SG_INF)
   OR (fSurgeP0 <= DL_SG_EPS) OR (fSurgeK < 0.0) THEN
    fMarginPct := 0.0;                // 裕度确定值零出口 / Deterministic zero margin
    eLevel     := E_DL_SurgeLevel.eNormal; // 参数不可信分级回正常（联锁侧另判）/ Level back to normal, interlock judged elsewhere
    uErrCode   := 16#0002_3921;       // 故障级：喘振线参数非法 / Fault: illegal surge line parameters
    bError     := TRUE;               // 置故障标志（R45 配对）/ Raise the fault flag, R45 pairing
    bValid     := FALSE;              // 输出不可用 / Outputs unusable
    RETURN;                           // 结构早退 / early exit
END_IF

// ---- 段 4｜工况点输入防御：非有限 → 信息级保持现状（分级冻结）----
IF (fFlowAct <> fFlowAct) OR (ABS(fFlowAct) > DL_SG_INF)
   OR (fPressAct <> fPressAct) OR (ABS(fPressAct) > DL_SG_INF) THEN
    uErrCode := 16#0002_3922;         // 信息级：工况点非有限 / Info: non-finite operating point
    bValid   := FALSE;                // 输出不可用（bTrip 锁存语义不变）/ Outputs unusable, trip latch semantics unchanged
    RETURN;                           // 结构早退（分级冻结不重算）/ early exit, level frozen
END_IF

// ---- 段 5｜裕度主体：线性喘振线取值 → 差值比；分母先过正域闸 ----
fPSurge := fSurgeP0 - fSurgeK * fFlowAct; // 喘振线压力 [Pa] / Surge line pressure [Pa]
IF fPSurge <= DL_SG_EPS THEN
    fPSurge := DL_SG_EPS;             // 深越线分母钳容差（防负/零除）/ Deep-beyond-line denominator clamped
END_IF
fMarginPct := (fPSurge - fPressAct) / fPSurge * DL_SG_PCT100; // 裕度 [百分数] / Margin [percent]

// ---- 段 6｜分级装配：裕度先判跳机带再判预警带（两级次序不可反）----
IF (fMarginPct <= fTripMargin) OR (fMarginPct < 0.0) THEN
    bInTripBand := TRUE;              // 跳机带或越线声明 / Trip band or beyond the line
ELSIF fMarginPct <= fWarnMargin THEN
    bInWarnBand := TRUE;              // 预警带声明 / Warning band
END_IF

// ---- 段 7｜锁存与确认：bTrip 锁存至复位沿/撤使能；去抖确认后才置声明 ----
IF trigReset.Q OR (NOT bEn) THEN
    bTrip := FALSE;                   // 锁存解除（复位沿或撤使能，头注释声明的清除沿）/ Latch released on reset edge or disable
END_IF
IF tonTrip.Q THEN
    bTrip := TRUE;                    // 跳机去抖确认置位 / Trip confirmed by debounce
END_IF
bWarn := tonWarn.Q AND NOT bTrip;     // 预警确认（跳机优先压制预警）/ Warning confirmed, suppressed by trip

// ---- 段 8｜分级状态机（CASE 带 ELSE；非法值兜底归 eTrip 安全侧）----
CASE eLevel OF
    E_DL_SurgeLevel.eNormal:          // 正常相：可升预警或跳机
        IF bTrip THEN
            eLevel := E_DL_SurgeLevel.eTrip;  // 升跳机 / Rise to trip
        ELSIF bWarn THEN
            eLevel := E_DL_SurgeLevel.eWarn;  // 升预警 / Rise to warning
            uErrCode := 16#0002_3920;         // 信息级：裕度进入预警带 / Info: margin in the warning band
        END_IF

    E_DL_SurgeLevel.eWarn:            // 预警相：可升跳机或降正常
        IF bTrip THEN
            eLevel := E_DL_SurgeLevel.eTrip;  // 升跳机 / Rise to trip
        ELSIF NOT bWarn THEN
            eLevel := E_DL_SurgeLevel.eNormal; // 降正常 / Fall back to normal
        ELSE
            uErrCode := 16#0002_3920;         // 预警保持期内信息级重算 / Info code recomputed while warning holds
        END_IF

    E_DL_SurgeLevel.eTrip:            // 跳机相：锁存，仅锁存解除后可降级
        IF NOT bTrip THEN             // 锁存已解除（复位沿/撤使能）
            IF bWarn THEN
                eLevel := E_DL_SurgeLevel.eWarn;  // 降预警 / Fall to warning
            ELSE
                eLevel := E_DL_SurgeLevel.eNormal; // 降正常 / Fall to normal
            END_IF
        END_IF

    ELSE                              // 非法分级兜底（R21：CASE 必带 ELSE）
        eLevel := E_DL_SurgeLevel.eTrip; // 拦截非法值归跳机（安全侧）/ Catch illegal value to trip, safe side
END_CASE

bValid := TRUE;                       // 全部防御通过：输出可用 / Outputs usable
END_FUNCTION_BLOCK

(* ---- FB_DL_FeedforwardComp.st ---- *)
(*==============================================================================
 * 组件名称 (Component)  : FB_DL_FeedforwardComp
 * 所属子库 (Sublibrary) : DL_Algo
 * 当前版本 (Version)    : 1.0.1
 * 兼容性   (Platform)   : CODESYS 3.5 / TwinCAT 3 / 汇川 InoProShop / Machine Expert
 *                         仅依赖纯 IEC 61131-3 数学运算，零库依赖，零厂商方言
 * 功能描述 (Function)   : 静态 + 动态前馈补偿器。对可测扰动量做前馈：静态增益
 *                         项即时响应 + 一阶惯性 / 超前滞后动态整形 + 可选纯滞后
 *                         （固定 10 槽延时队列），输出叠加到 PID 反馈通道，提升
 *                         抗负载扰动速度。现场用途：配料设定突变、蒸汽压力波动
 *                         的前馈补偿。
 * 开源溯源 (Origin)     : 原创实现。超前滞后 / 纯滞后补偿功能分类与参数域参考
 *                         过程控制经典文献（lead-lag and dead-time feedforward）
 *                         的公开语义描述，未复制任何厂商源码，clean-room 重写。
 * 本文件内含       : TYPE  E_DL_FfState（配套枚举，归属 DL_Algo）
 *                    FB    FB_DL_FeedforwardComp
 * 依赖     (Depends)    : 无 DL_ 内部依赖；Standard.library 无实例依赖
 * 红线自检 (Redline)    : R1 ✓ 零全局变量表与外部变量引用 ｜ R2 ✓ 零物理 IO 地址直写
 *                         R3 ✓ 纯 IEC 61131-3 ｜ R4 ✓ 防除零+钳位+数组边界防御
 *                         R5 ✓ 全变量中英双语同行注释 ｜ R6 ✓ 四态 ENUM+CASE+ELSE
 *                         R7 ✓ 本块无定时器 / 边沿实例（无可刷新项，天然合规）
 * 修订历史 (Revision)   :
 *   2026-11-15  v1.0.0  首版入库 · Round 04 · Level 1 DL_Algo
 *   2026-11-15  v1.0.1  阶段五终审精修：tLagTime=T#0S 为规格合法直通口径，
 *                       不再误置 0002_0401 故障码
 * 验收向量 (Acceptance) :
 *   V1 纯静态：tLead=tLag=tDelay=T#0S, fFfGain=2, 扰动=10 → fFfOut=20
 *   V2 惯性收敛：tLag=T#1S, 恒扰动 10 → fDynPart 单调趋近扰动值
 *   V3 滞后：tDelay=T#300MS, 扰动阶跃 → 输出滞后 3 拍后出现
 *   V4 跟踪：bTrack 置位 → fFfOut 立即等于钳位后的 fTrackValue
 *   V5 队列截断：tDelay 折算深度超 10 → nDelaySteps=10 且码 0002_0402
 *   V6 非有限值：扰动写非法浮点 → 输出保持上一拍且码 0002_0004
 *============================================================================*)

(*-----------------------------------------------------------------------------
 * 枚举: E_DL_FfState（归属 DL_Algo，与 FB_DL_FeedforwardComp 同文件）
 * 含义: 前馈补偿离散状态。数值步长留空位便于后续插态而不破坏已有工程。
 *----------------------------------------------------------------------------*)
TYPE E_DL_FfState :
(
    eIdle    := 0,    // 使能关：输出回下限，队列冻结 / Idle: enable off, output at low limit
    eStatic  := 10,   // 仅静态：超前滞后与滞后队列全关 / Static only: lead-lag and delay queue off
    eDynamic := 20,   // 动态：惯性 / 超前 / 滞后环节至少一项使能 / Dynamic: at least one shaping element active
    eFault   := 99    // 故障兜底态：非法状态进入，输出安全值 / Fault fallback: illegal state, safe output
);
END_TYPE

(*==============================================================================
 * 功能块: FB_DL_FeedforwardComp
 * 调用约定: 每个扫描周期无条件调用一次；滞后队列每拍必须持续写入。
 * 无状态泄漏: 全部状态驻留于实例私有 VAR，零全局引用，可多实例并行。
 * 工程披露: 滞后队列为固定 10 槽环形缓冲，深度按 tDelayTime/tSampleTime 向下
 *           取整折算，超出上限截断并置码，不做动态扩容。
 *============================================================================*)
FUNCTION_BLOCK FB_DL_FeedforwardComp
VAR_INPUT
    bEnable     : BOOL := FALSE;      // 总使能，FALSE 时输出回下限 / Master enable, FALSE drives output to low limit
    fDisturbance: REAL := 0.0;        // 扰动量 [EU]，可测负载信号 / Measured disturbance in engineering units
    fFfGain     : REAL := 1.0;        // 前馈增益 [1] / Feedforward gain, dimensionless
    tLeadTime   : TIME := T#0S;       // 超前时间 [s]，T#0S = 纯静态 / Lead time [s], T#0S = static only
    tLagTime    : TIME := T#0S;       // 惯性时间 [s]，T#0S = 直通 / Lag time [s], T#0S = pass-through
    tDelayTime  : TIME := T#0S;       // 纯滞后时间 [s]，T#0S = 无滞后队列 / Dead time [s], T#0S = no queue
    rOutMin     : REAL := -100.0;     // 输出下限 [%] / Output lower limit in percent
    rOutMax     : REAL := 100.0;      // 输出上限 [%] / Output upper limit in percent
    tSampleTime : TIME := T#100MS;    // 采样周期 [s] / Sample period in seconds
    bTrack      : BOOL := FALSE;      // 跟踪使能，TRUE 时输出立即跟随跟踪值 / Track enable, output follows track value
    fTrackValue : REAL := 0.0;        // 跟踪值 [%]，用于无扰投切 / Track value in percent
END_VAR
VAR_OUTPUT
    fFfOut      : REAL;               // 前馈输出 [%] / Feedforward output in percent
    fStaticPart : REAL;               // 静态分量 [%]，诊断 / Static component, diagnostics
    fDynPart    : REAL;               // 动态分量 [%]，诊断 / Dynamic component, diagnostics
    bError      : BOOL;               // 故障标志 / Fault flag
    uErrorId    : UDINT;              // 故障码，0 = 无故障 / Error code, 0 = no error
END_VAR
VAR
    fDyn        : REAL;               // 惯性环节状态 [EU] / Inertia element state
    fDynPrev    : REAL;               // 上一拍惯性状态 [EU]，诊断 / Previous inertia state, diagnostics
    afDelayBuf  : ARRAY[0..9] OF REAL;// 滞后队列 [EU]，固定 10 槽环形 / Delay queue, fixed 10-slot ring
    nDelaySteps : INT;                // 队列深度 = tDelayTime/tSampleTime [拍] / Queue depth in cycles
    nWriteIdx   : INT;                // 环形队列写指针 [0..9] / Ring buffer write index
    eState      : E_DL_FfState;       // 主状态机当前状态 / Current state of the state machine
    bInit       : BOOL := FALSE;      // 首扫初始化标志 / First-scan init flag
    fDt         : REAL;               // 生效采样周期 [s] / Effective sample period in seconds
    fLimLow     : REAL;               // 修复后的输出下限 [%] / Repaired output lower limit
    fLimHigh    : REAL;               // 修复后的输出上限 [%] / Repaired output upper limit
    fLeadFactor : REAL;               // 超前因子 [1] / Lead factor, dimensionless
    fDelayed    : REAL;               // 滞后队列读出值 [EU] / Delayed value read from queue
    fFfRaw      : REAL;               // 限幅前的原始前馈输出 [%] / Raw feedforward output before clamp
    nReadIdx    : INT;                // 环形队列读指针 [0..9] / Ring buffer read index
    nDepthRaw   : INT;                // 折算的原始队列深度 [拍] / Raw computed queue depth in cycles
    bNonFinite  : BOOL;               // 本拍输入非有限值标志 / Non-finite input flag of this cycle
END_VAR
VAR CONSTANT
    DL_FF_DELAY_MAX : INT := 10;      // 滞后队列深度上限 [槽] / Delay queue depth ceiling in slots
END_VAR

(*------------------------------------------------------------------------------
 * 段 1｜参数钳位与公共防御（不中断扫描）
 *      Parameter clamping and common defenses, never stops the scan
 *-----------------------------------------------------------------------------*)
bError   := FALSE;                    // 每拍重算故障标志 / Recompute fault flag every cycle
uErrorId := 16#0002_0000;             // 每拍重算故障码 / Recompute error code every cycle
bNonFinite := FALSE;                  // 非有限值标志每拍重算 / Non-finite flag recomputed every cycle

IF tSampleTime < T#10MS THEN
    fDt := 0.01;                      // 采样周期非法钳位为 0.01 s / Illegal sample period clamped to 0.01 s
    uErrorId := 16#0002_0002;         // 公共码：采样周期已钳位 / Common code: sample period clamped
ELSE
    fDt := TIME_TO_REAL(tSampleTime) / 1000.0;  // 采样周期换算为秒 [s] / Sample period in seconds
END_IF

IF rOutMin > rOutMax THEN
    fLimLow  := rOutMax;              // 上下限对调修复 / Swapped repair of limits
    fLimHigh := rOutMin;              // 上下限对调修复 / Swapped repair of limits
    uErrorId := 16#0002_0001;         // 公共码：参数越界已钳位 / Common code: parameter clamped
ELSE
    fLimLow  := rOutMin;              // 合法下限直通 / Valid low limit passed
    fLimHigh := rOutMax;              // 合法上限直通 / Valid high limit passed
END_IF

(* 输入非有限值防御：扰动或跟踪值非法即拒绝本拍更新 *)
(* Non-finite defense: reject this cycle if disturbance or track value invalid *)
IF (fDisturbance <> fDisturbance) OR (ABS(fDisturbance) > 1.0E30)
   OR (fTrackValue <> fTrackValue) OR (ABS(fTrackValue) > 1.0E30) THEN
    bNonFinite := TRUE;               // 置非有限值标志 / Set non-finite flag
    bError   := TRUE;                 // 置故障标志 / Set fault flag
    uErrorId := 16#0002_0004;         // 公共码：输入非有限值已拒绝 / Common code: non-finite rejected
END_IF

(*------------------------------------------------------------------------------
 * 段 2｜队列深度折算：tDelayTime/tSampleTime 向下取整，超上限截断置码
 *      Queue depth derivation: floor division, truncated at ceiling with code
 *-----------------------------------------------------------------------------*)
nDepthRaw := REAL_TO_INT(TRUNC(TIME_TO_REAL(tDelayTime) / 1000.0 / fDt));  // 原始深度 [拍] / Raw depth in cycles
IF nDepthRaw > DL_FF_DELAY_MAX THEN
    nDelaySteps := DL_FF_DELAY_MAX;   // 深度截断至上限 / Depth truncated to ceiling
    uErrorId := 16#0002_0402;         // 组件码：滞后队列深度超上限已截断 / Code: queue depth truncated
ELSIF nDepthRaw < 0 THEN
    nDelaySteps := 0;                 // 负深度防御为 0 / Negative depth defended to zero
ELSE
    nDelaySteps := nDepthRaw;         // 合法深度直通 / Valid depth passed
END_IF

(*------------------------------------------------------------------------------
 * 段 3｜使能与跟踪早退：保持上一拍输出，队列冻结
 *      Early exit on disable or track: hold output, queue frozen
 *-----------------------------------------------------------------------------*)
IF NOT bEnable THEN
    eState    := eIdle;               // 强制回空闲态 / Force idle state
    fFfOut    := fLimLow;             // 输出回下限 / Output to low limit
    fStaticPart := 0.0;               // 静态分量清零 / Static component cleared
    fDynPart  := 0.0;                 // 动态分量清零 / Dynamic component cleared
    RETURN;                           // 本拍结束 / End of this cycle
END_IF

IF bNonFinite THEN
    RETURN;                           // 保持上一拍输出与状态 / Hold previous output and state
END_IF

IF bTrack OR (NOT bInit) THEN
    (* 跟踪回投 / 首扫初始化：输出立即跟随，惯性状态与队列同步，投切无扰 *)
    (* Track / first-scan init: output follows, inertia state and queue in sync *)
    IF bTrack THEN
        fFfOut := LIMIT(fLimLow, fTrackValue, fLimHigh);          // 输出钳位跟随 / Clamped tracking output
    ELSE
        fFfOut := fLimLow;            // 首扫输出回下限 / First-scan output to low limit
    END_IF
    fDyn        := fDisturbance;      // 惯性状态同步 / Inertia state synchronized
    fDynPrev    := fDisturbance;      // 上拍惯性状态同步 / Previous state synchronized
    FOR nReadIdx := 0 TO DL_FF_DELAY_MAX - 1 DO
        afDelayBuf[nReadIdx] := fDisturbance;                     // 队列全槽预填 / Prefill all queue slots
    END_FOR
    nWriteIdx   := 0;                 // 写指针归零 / Write index reset
    bInit       := TRUE;              // 置首扫完成标志 / Set first-scan done flag
    fStaticPart := 0.0;               // 静态分量清零 / Static component cleared
    fDynPart    := 0.0;               // 动态分量清零 / Dynamic component cleared
    RETURN;                           // 本拍结束 / End of this cycle
END_IF

(*------------------------------------------------------------------------------
 * 段 4｜前馈计算：静态项 + 动态项（惯性 / 超前）+ 纯滞后队列
 *      Feedforward computation: static term plus dynamic and dead-time terms
 *-----------------------------------------------------------------------------*)
fStaticPart := fFfGain * fDisturbance;                            // 静态项即时响应 [%] / Static term, instant response

(* 状态派生：任一动态环节使能即进动态态 *)
(* State derivation: any shaping element active means dynamic state *)
IF (tLeadTime = T#0S) AND (tLagTime = T#0S) AND (tDelayTime = T#0S) THEN
    eState := eStatic;                // 仅静态 / Static only
ELSE
    eState := eDynamic;               // 动态使能 / Dynamic active
END_IF

IF eState = eDynamic THEN
    (* 动态项：一阶超前 / 惯性离散差分，tLagTime 小于一拍时按一拍直通 *)
    (* Dynamic term: first-order lead/lag recursion, sub-cycle lag treated as one-cycle *)
    fLeadFactor := 1.0 + TIME_TO_REAL(tLeadTime) / 1000.0 / fDt;  // 超前因子 [1] / Lead factor
    IF tLeadTime < T#0S THEN
        fLeadFactor := 1.0;           // 负超前防御为 1（关闭超前） / Negative lead defended to 1
        uErrorId := 16#0002_0401;     // 组件码：动态时间非法已钳位 / Code: dynamic time clamped
    END_IF
    IF tLagTime <= T#0S THEN
        fDyn := fDisturbance;         // T#0S = 直通，规格合法口径不置故障码 / T#0S = pass-through, legal per spec, no error code
    ELSE
        fDyn := fDyn + (fLeadFactor * fDisturbance - fDyn) * fDt
                    / MAX(TIME_TO_REAL(tLagTime) / 1000.0, fDt);  // 惯性递推 / Inertia recursion
    END_IF
    fDynPrev := fDyn;                 // 上拍惯性状态记录 / Record previous inertia state

    (* 纯滞后队列：先写入当前值，再按深度回读，指针经取模保证不越界 *)
    (* Dead-time queue: write current value first, read back by depth, modulo safe *)
    afDelayBuf[nWriteIdx] := fDisturbance;                        // 当前扰动入队 / Enqueue current disturbance
    nReadIdx := (nWriteIdx - nDelaySteps + DL_FF_DELAY_MAX) MOD DL_FF_DELAY_MAX;  // 读指针 / Read index
    nReadIdx := LIMIT(0, nReadIdx, DL_FF_DELAY_MAX - 1);          // 读指针防御钳位 / Defensive index clamp
    fDelayed := afDelayBuf[nReadIdx];                             // 滞后读出 [EU] / Delayed readout
    nWriteIdx := (nWriteIdx + 1) MOD DL_FF_DELAY_MAX;             // 写指针推进 / Advance write index
    fDynPart := fFfGain * (fDyn - fDelayed);                      // 动态分量 [%] / Dynamic component
ELSE
    fDelayed  := fDisturbance;        // 静态模式无滞后 / Static mode has no delay
    fDynPart  := 0.0;                 // 动态分量清零 / Dynamic component cleared
    fDynPrev  := fDisturbance;        // 惯性状态直通同步 / Inertia state pass-through
END_IF

fFfRaw := fStaticPart + fDynPart;     // 原始前馈合成 [%] / Raw feedforward composition
fFfOut := LIMIT(fLimLow, fFfRaw, fLimHigh);                       // 输出限幅 / Output clamping

(*------------------------------------------------------------------------------
 * 段 5｜主状态机收口（红线 R6）：CASE 覆盖 + ELSE 兜底
 *      State machine closure: CASE coverage with mandatory ELSE fallback
 *-----------------------------------------------------------------------------*)
CASE eState OF
    eIdle:    ;                        // 空闲态已在早退段处理 / Idle handled in early exit
    eStatic:  ;                        // 静态态输出已合成 / Static output composed
    eDynamic: ;                        // 动动态输出已合成 / Dynamic output composed
    eFault:   ;                        // 故障态占位（参数故障不锁存控制） / Fault placeholder
    ELSE
        (* 非法状态拦截：一律进故障兜底并置码 *)
        (* Illegal state interception: force fault fallback with code *)
        eState   := eFault;            // 进故障态 / Enter fault state
        bError   := TRUE;              // 置故障标志 / Set fault flag
        uErrorId := 16#0002_0005;      // 非法状态兜底码 / Illegal state fallback code
        fFfOut   := fLimLow;           // 安全输出 / Safe output
END_CASE;
END_FUNCTION_BLOCK
